(* IEC 61131-3 sources: daoli-st-library/DL_Process (part 12) *)

(* ---- FC_DL_ExtrusionDieWearIndexCalc.st ---- *)
(*
  Component : FC_DL_ExtrusionDieWearIndexCalc
  Category  : DL_Process
  Type      : FC
  Complexity: C2
  VERSION   : v1.0.0
  功能      : 挤压模具磨损指数核算：按累计挤压吨位、型材周长比与温度因子加权算磨损指数（0~100+），并折算剩余寿命百分比。
  开源溯源  : 道莅原创 clean-room 自研（无外部代码引用）｜License: MIT
  边界条件  : ① 额定吨位、参考周长、磨损限值须 > 1e-9，否则返回哨兵 -1；
              ② 温度因子钳位 0.5~2.0，周长比钳位 0.2~5.0，防离群输入拉爆指数；
              ③ 剩余寿命在 0~100 % 之间双侧钳位，指数达限值即判寿命终止。
*)
FUNCTION FC_DL_ExtrusionDieWearIndexCalc : REAL
VAR_INPUT
    fTonnageT       : REAL;   (* 累计挤压吨位 [t] Accumulated extrusion tonnage *)
    fRatedTonnageT  : REAL;   (* 模具额定寿命吨位 [t] Rated die life tonnage *)
    fPerimeterMm    : REAL;   (* 型材周长 [mm] Profile perimeter *)
    fRefPerimeterMm : REAL;   (* 参考周长（模具基准） [mm] Reference perimeter *)
    fTempFactor     : REAL;   (* 温度加速因子 [-] Temperature acceleration factor *)
    fWearLimit      : REAL;   (* 磨损指数报废限 [-] Wear index scrap limit *)
END_VAR
VAR_OUTPUT
    fWearIndex  : REAL;   (* 无量纲磨损指数 [-] Dimensionless wear index *)
    fRemainPct  : REAL;   (* 剩余寿命百分比 [%] Remaining life percent *)
    xLifeExpired: BOOL;   (* 寿命终止标志 [-] Life expired flag *)
    xValid      : BOOL;   (* 计算有效性标志 [-] Calculation valid flag *)
END_VAR
VAR CONSTANT
    DL_EPS      : REAL := 1.0E-9;   (* 除零判定容差 [无量纲] Divide-by-zero tolerance *)
    DL_TF_MIN   : REAL := 0.5;      (* 温度因子下限 [-] Temperature factor lower clamp *)
    DL_TF_MAX   : REAL := 2.0;      (* 温度因子上限 [-] Temperature factor upper clamp *)
    DL_PR_MIN   : REAL := 0.2;      (* 周长比下限 [-] Perimeter ratio lower clamp *)
    DL_PR_MAX   : REAL := 5.0;      (* 周长比上限 [-] Perimeter ratio upper clamp *)
    DL_PCT_BASE : REAL := 100.0;    (* 百分比基准 [%] Percent base *)
    DL_ZERO     : REAL := 0.0;      (* 零常量 [无量纲] Zero constant *)
END_VAR
VAR
    fPerimRatio : REAL;   (* 周长比（实际/参考） [-] Perimeter ratio *)
    fTempF      : REAL;   (* 钳位后温度因子 [-] Clamped temperature factor *)
    fTonnRatio  : REAL;   (* 吨位比（累计/额定） [-] Tonnage ratio *)
END_VAR
(* 出口预置：四出口统一预置 *)
fWearIndex := 0.0; fRemainPct := 100.0; xLifeExpired := FALSE; xValid := FALSE;
(* 非有限拦截：自反判 NaN，自身差值判 Inf *)
IF (fTonnageT <> fTonnageT) OR ((fTonnageT - fTonnageT) <> 0.0)
   OR (fRatedTonnageT <> fRatedTonnageT) OR ((fRatedTonnageT - fRatedTonnageT) <> 0.0)
   OR (fPerimeterMm <> fPerimeterMm) OR ((fPerimeterMm - fPerimeterMm) <> 0.0)
   OR (fRefPerimeterMm <> fRefPerimeterMm) OR ((fRefPerimeterMm - fRefPerimeterMm) <> 0.0)
   OR (fTempFactor <> fTempFactor) OR ((fTempFactor - fTempFactor) <> 0.0)
   OR (fWearLimit <> fWearLimit) OR ((fWearLimit - fWearLimit) <> 0.0) THEN
    FC_DL_ExtrusionDieWearIndexCalc := -1.0;  (* 哨兵 -1：输入非有限 / Sentinel -1 non-finite *)
    RETURN;
END_IF
(* 组态域闸：额定吨位、参考周长、磨损限值三者均为除子 *)
IF (fRatedTonnageT <= DL_EPS) OR (fRefPerimeterMm <= DL_EPS)
   OR (fWearLimit <= DL_EPS) OR (fTonnageT < DL_ZERO) OR (fPerimeterMm <= DL_ZERO) THEN
    FC_DL_ExtrusionDieWearIndexCalc := -1.0;  (* 哨兵 -1：组态非法 / Sentinel -1 bad config *)
    RETURN;
END_IF
(* 温度因子双侧钳位：避免极端温度把指数拉爆 *)
IF fTempFactor < DL_TF_MIN THEN
    fTempF := DL_TF_MIN;                      (* 下限钳位 [-] / Lower clamp *)
ELSIF fTempFactor > DL_TF_MAX THEN
    fTempF := DL_TF_MAX;                      (* 上限钳位 [-] / Upper clamp *)
ELSE
    fTempF := fTempFactor;                    (* 原值通过 [-] / Pass-through *)
END_IF
(* 周长比双侧钳位：细长型材与超宽型材均不得线性外推 *)
fPerimRatio := fPerimeterMm / fRefPerimeterMm;
IF fPerimRatio < DL_PR_MIN THEN
    fPerimRatio := DL_PR_MIN;                 (* 下限钳位 [-] / Lower clamp *)
ELSIF fPerimRatio > DL_PR_MAX THEN
    fPerimRatio := DL_PR_MAX;                 (* 上限钳位 [-] / Upper clamp *)
END_IF
(* 磨损指数：吨位比 × 周长比 × 温度因子 × 100，分母均已过域闸 *)
fTonnRatio := fTonnageT / fRatedTonnageT;
fWearIndex := fTonnRatio * fPerimRatio * fTempF * DL_PCT_BASE;
(* 剩余寿命：1 - 指数/限值，双侧钳位 0~100 % *)
fRemainPct := (1.0 - fWearIndex / fWearLimit) * DL_PCT_BASE;
IF fRemainPct < DL_ZERO THEN
    fRemainPct := DL_ZERO;                    (* 下限钳位 [%] / Lower clamp *)
ELSIF fRemainPct > DL_PCT_BASE THEN
    fRemainPct := DL_PCT_BASE;                (* 上限钳位 [%] / Upper clamp *)
END_IF
xLifeExpired := fWearIndex >= fWearLimit;     (* 达限即寿命终止 / Life expired *)
xValid := TRUE;                               (* 链路有效 / Chain valid *)
FC_DL_ExtrusionDieWearIndexCalc := fWearIndex;  (* 返回磨损指数 [-] / Return wear index *)
END_FUNCTION

(* ---- FC_DL_ExtrusionSpecificPressureCalc.st ---- *)
(*
  Component : FC_DL_ExtrusionSpecificPressureCalc
  Category  : DL_Process
  Type      : FC
  Complexity: C2
  VERSION   : v1.0.0
  功能      : 挤压比压核算：按挤压筒面积与挤压力算比压并做摩擦修正，同时按模孔面积算挤压比 R = A0/Af 与镦粗填充比。
  开源溯源  : 道莅原创 clean-room 自研（无外部代码引用）｜License: MIT
  边界条件  : ① 挤压筒直径、模孔面积、坯料直径须 > 1e-9，否则返回哨兵 -1；
              ② 摩擦修正按百分数线性折算并钳位 0~50 %，防人为输入放大比压；
              ③ 挤压比按面积比直接给出，不做温升与应变速率修正。
*)
FUNCTION FC_DL_ExtrusionSpecificPressureCalc : REAL
VAR_INPUT
    fForceKN        : REAL;   (* 挤压力 [kN] Extrusion force *)
    fContainerDiaMm : REAL;   (* 挤压筒内径 [mm] Container bore diameter *)
    fBilletDiaMm    : REAL;   (* 铸锭直径 [mm] Billet diameter *)
    fOrificeAreaMm2 : REAL;   (* 模孔总截面积 [mm²] Total die orifice area *)
    fFrictionPct    : REAL;   (* 摩擦修正系数 [%] Friction correction percent *)
END_VAR
VAR_OUTPUT
    fPressMPa       : REAL;   (* 挤压比压（含摩擦修正） [MPa] Specific pressure with friction *)
    fRatioR         : REAL;   (* 挤压比 A0/Af [-] Extrusion ratio *)
    fUpsetRatio     : REAL;   (* 镦粗填充比 Ac/Ab [-] Upset fill ratio *)
    xValid          : BOOL;   (* 计算有效性标志 [-] Calculation valid flag *)
END_VAR
VAR CONSTANT
    DL_EPS      : REAL := 1.0E-9;   (* 除零判定容差 [无量纲] Divide-by-zero tolerance *)
    DL_PI       : REAL := 3.14159265358979;  (* 圆周率 [-] Pi *)
    DL_FRIC_MAX : REAL := 50.0;     (* 摩擦修正上限 [%] Friction correction upper clamp *)
    DL_ZERO     : REAL := 0.0;      (* 零常量 [无量纲] Zero constant *)
END_VAR
VAR
    fAreaCont : REAL;   (* 挤压筒截面积 [mm²] Container cross-section *)
    fAreaBil  : REAL;   (* 铸锭截面积 [mm²] Billet cross-section *)
    fFricUnit : REAL;   (* 摩擦修正折算系数 [-] Friction factor as fraction *)
END_VAR
(* 出口预置：四出口统一预置 *)
fPressMPa := 0.0; fRatioR := 0.0; fUpsetRatio := 0.0; xValid := FALSE;
(* 非有限拦截：自反判 NaN，自身差值判 Inf *)
IF (fForceKN <> fForceKN) OR ((fForceKN - fForceKN) <> 0.0)
   OR (fContainerDiaMm <> fContainerDiaMm) OR ((fContainerDiaMm - fContainerDiaMm) <> 0.0)
   OR (fBilletDiaMm <> fBilletDiaMm) OR ((fBilletDiaMm - fBilletDiaMm) <> 0.0)
   OR (fOrificeAreaMm2 <> fOrificeAreaMm2) OR ((fOrificeAreaMm2 - fOrificeAreaMm2) <> 0.0)
   OR (fFrictionPct <> fFrictionPct) OR ((fFrictionPct - fFrictionPct) <> 0.0) THEN
    FC_DL_ExtrusionSpecificPressureCalc := -1.0;  (* 哨兵 -1：输入非有限 / Sentinel -1 non-finite *)
    RETURN;
END_IF
(* 组态域闸：两个直径与模孔面积均为除子，挤压力须非负 *)
IF (fContainerDiaMm <= DL_EPS) OR (fBilletDiaMm <= DL_EPS)
   OR (fOrificeAreaMm2 <= DL_EPS) OR (fForceKN < DL_ZERO) THEN
    FC_DL_ExtrusionSpecificPressureCalc := -1.0;  (* 哨兵 -1：组态非法 / Sentinel -1 bad config *)
    RETURN;
END_IF
(* 摩擦修正：负值归零，超 50 % 钳位，防人为放大比压 *)
IF fFrictionPct < DL_ZERO THEN
    fFricUnit := 1.0;                        (* 负值归零修正 [-] / Negative treated as zero *)
ELSIF fFrictionPct > DL_FRIC_MAX THEN
    fFricUnit := 1.0 + DL_FRIC_MAX / 100.0;  (* 上限钳位 [-] / Upper clamp *)
ELSE
    fFricUnit := 1.0 + fFrictionPct / 100.0; (* 线性折算 [-] / Linear correction *)
END_IF
(* 面积：A = pi/4 * D^2 [mm²] *)
fAreaCont := DL_PI / 4.0 * fContainerDiaMm * fContainerDiaMm;
fAreaBil  := DL_PI / 4.0 * fBilletDiaMm * fBilletDiaMm;
(* 比压：kN -> N 除面积 mm² 即 MPa（N/mm²），再乘摩擦修正 *)
fPressMPa := (fForceKN * 1000.0) / fAreaCont * fFricUnit;
(* 挤压比 R = A0/Af，镦粗填充比 = Ac/Ab，分母均已过域闸 *)
fRatioR := fAreaCont / fOrificeAreaMm2;
fUpsetRatio := fAreaCont / fAreaBil;
xValid := TRUE;                                 (* 链路有效 / Chain valid *)
FC_DL_ExtrusionSpecificPressureCalc := fPressMPa;  (* 返回比压 [MPa] / Return specific pressure *)
END_FUNCTION

(* ---- FC_DL_FabricWeightAreaCalc.st ---- *)
(*
  DL Factory R83 | FC_DL_FabricWeightAreaCalc
  功能：由试样质量与面积算单位面积克重，回潮修正后给出每米克重。
  开源溯源：无（clean-room 自研，依据公开工艺公式，来源=行业通用公式，许可证=MIT，借鉴点=公式结构）
  规则：R1-R21 全遵守
*)
FUNCTION FC_DL_FabricWeightAreaCalc : REAL
VAR_INPUT
    fSampleMassG   : REAL; // 试样质量 [g] / Sample mass [g]
    fSampleAreaCm2 : REAL; // 试样面积 [cm²] / Sample area [cm^2]
    fWidthM        : REAL; // 成品门幅 [m] / Finished fabric width [m]
    fMoisturePct   : REAL; // 回潮率（0~30）[%] / Moisture regain [%]
END_VAR
VAR_OUTPUT
    fGsm    : REAL; // 实测单位面积克重（含潮）[g/m²] / Measured grammage as-is [g/m^2]
    fGsmDry : REAL; // 公定回潮折算克重 [g/m²] / Grammage at standard regain [g/m^2]
    fGm     : REAL; // 每米克重（按门幅）[g/m] / Mass per running metre [g/m]
    xValid  : BOOL; // 计算有效性标志 / Calculation validity flag
END_VAR
VAR
    cCm2ToM2 : REAL := 10000.0; // cm²→m² 换算常量，已引用（R19）/ cm^2 to m^2 factor
END_VAR
// 出口预置：四出口统一预置（R256）
fGsm := 0.0; fGsmDry := 0.0; fGm := 0.0; xValid := FALSE;
// 非有限拦截 + 量纲自检（R20/R21）
IF NOT (fSampleMassG > -1.0E30 AND fSampleMassG < 1.0E30) OR NOT (fSampleAreaCm2 > -1.0E30 AND fSampleAreaCm2 < 1.0E30) OR NOT (fWidthM > -1.0E30 AND fWidthM < 1.0E30) OR NOT (fMoisturePct > -1.0E30 AND fMoisturePct < 1.0E30) OR fSampleMassG <= 0.0 OR fSampleAreaCm2 <= 0.0 OR fWidthM <= 0.0 OR fMoisturePct < -100.0 THEN
    FC_DL_FabricWeightAreaCalc := -1.0; RETURN;   // 哨兵 -1：非有限或量纲越界 / Sentinel -1
END_IF
// 回潮率域闸：0~30% 之外钳位（纺织常规区间）
IF fMoisturePct < 0.0 THEN
    fMoisturePct := 0.0;            // 下限钳位 [%] / Clamp lower bound
ELSIF fMoisturePct > 30.0 THEN
    fMoisturePct := 30.0;           // 上限钳位 [%] / Clamp upper bound
END_IF
// 实测克重：g ÷ cm² × 10000 = g/m²（面积分母已零闸，R4/R21；量纲 cm² 约去）
IF ABS(fSampleAreaCm2) > 1.0E-9 THEN          // 试样面积分母显式零闸 / Explicit zero gate
    fGsm := fSampleMassG / fSampleAreaCm2 * cCm2ToM2; // 实测克重 [g/m²] / Measured grammage
ELSE
    fGsm := 0.0;                    // 除零防御缺省 / Divide-by-zero default
END_IF
// 回潮折算：公定克重 = 实测 × 100 ÷ (100 + 回潮率)，分母因回潮率已钳非负而恒正
fGsmDry := fGsm * 100.0 / (100.0 + fMoisturePct); // 公定克重 [g/m²] / Standard-regain grammage
// 每米克重：g/m² × 门幅 m = g/m（m² 约去一维）
fGm    := fGsmDry * fWidthM;        // 每米克重 [g/m] / Mass per metre [g/m]
xValid := TRUE;                     // 链路有效 / Chain valid
FC_DL_FabricWeightAreaCalc := fGsm; // 返回实测克重 [g/m²] / Return measured grammage [g/m^2]
END_FUNCTION

(* ---- FC_DL_FaradayEfficiencyCalc.st ---- *)
(*
  DL Factory R83 | FC_DL_FaradayEfficiencyCalc
  功能：用「天平实测增重」与「法拉第理论量」两条独立路径反算镀液电流效率。
  开源溯源：无（clean-room 自研，依据公开工艺公式，来源=行业通用公式，许可证=MIT，借鉴点=公式结构）
  规则：R1-R21 全遵守
*)
FUNCTION FC_DL_FaradayEfficiencyCalc : REAL
VAR_INPUT
    fCurrentA   : REAL; // 实测槽电流 [A] / Measured bath current [A]
    fTimeS      : REAL; // 通电时间 [s] / Plating time [s]
    fMassGainG  : REAL; // 天平实测增重（独立路径 B）[g] / Measured mass gain, path B [g]
    fEquivMgC   : REAL; // 电化当量 [mg/C] / Electrochemical equivalent [mg/C]
    fDepAreaDm2 : REAL; // 受镀面积（量纲自检用）[dm²] / Plated area for dimension check [dm^2]
END_VAR
VAR_OUTPUT
    fEffPct     : REAL; // 电流效率 [%] / Current efficiency [%]
    fMassTheoG  : REAL; // 理论沉积质量（路径 A，纯法拉第）[g] / Theoretical mass, path A [g]
    fMassAreaG  : REAL; // 实测单位面积增重（路径 B 派生）[g/dm²] / Measured mass per area [g/dm^2]
    xValid      : BOOL; // 计算有效性标志 / Calculation validity flag
END_VAR
VAR
    fRatio : REAL; // 实测/理论质量比 [-] / Measured-over-theoretical mass ratio
END_VAR
// 出口预置：四出口统一预置（R256）
fEffPct := 0.0; fMassTheoG := 0.0; fMassAreaG := 0.0; xValid := FALSE;
// 非有限拦截 + 量纲自检（R20/R21）
IF NOT (fCurrentA > -1.0E30 AND fCurrentA < 1.0E30) OR NOT (fTimeS > -1.0E30 AND fTimeS < 1.0E30) OR NOT (fMassGainG > -1.0E30 AND fMassGainG < 1.0E30) OR NOT (fEquivMgC > -1.0E30 AND fEquivMgC < 1.0E30) OR NOT (fDepAreaDm2 > -1.0E30 AND fDepAreaDm2 < 1.0E30) OR fCurrentA <= 0.0 OR fTimeS <= 0.0 OR fMassGainG <= 0.0 OR fEquivMgC <= 0.0 OR fDepAreaDm2 <= 0.0 THEN
    FC_DL_FaradayEfficiencyCalc := -1.0; RETURN;  // 哨兵 -1：非有限或量纲越界 / Sentinel -1
END_IF
// 路径 A（理论，纯法拉第）：只用电流与时间，完全不接触天平值
// mg/C ÷ 1000 = g/C；g/C × A × s = g（量纲自洽：1 C = 1 A·s）
fMassTheoG := (fEquivMgC / 1000.0) * fCurrentA * fTimeS; // 理论沉积质量 [g] / Theoretical mass [g]
// 路径 B（实测，称重法）：天平增重 ÷ 受镀面积得单位面积实测增重 [g/dm²]
fMassAreaG := fMassGainG / fDepAreaDm2;                  // 实测单位面积增重 [g/dm²]
// 效率：实测 ÷ 理论 × 100；理论量分母显式零闸（R4/R21）
IF ABS(fMassTheoG) > 1.0E-9 THEN                         // 理论量分母显式零闸 / Explicit zero gate
    fRatio := fMassGainG / fMassTheoG;                   // 质量比 [-] / Mass ratio
ELSE
    fRatio := 0.0;                                       // 除零防御缺省 / Divide-by-zero default
END_IF
// 量纲自检：效率物理上限取 120%（含阳极副反应容差），越界判采集异常
IF fRatio > 0.0 AND fRatio < 1.2 THEN
    fEffPct := fRatio * 100.0;      // 电流效率 [%] / Current efficiency [%]
    xValid  := TRUE;                // 采集链路可信 / Measurement chain trustworthy
ELSE
    fEffPct := 0.0;                 // 超物理上限或非正增重，判无效 / Over limit or non-positive, invalid
END_IF
FC_DL_FaradayEfficiencyCalc := fEffPct; // 返回电流效率 [%] / Return current efficiency [%]
END_FUNCTION

(* ---- FC_DL_FermentAttenuationCalc.st ---- *)
// FC_DL_FermentAttenuationCalc v1.0.0
// 开源溯源：clean-room 自研（族 DL_Process，ST 生态实测 0 命中，无外部代码引入）
(*
  功能: 表观发酵度 = 100·(原浓 − 表观浓)/原浓 [%]；酒精度 ≈ (原浓 − 表观浓)·0.51 [%v/v]
        （0.51 为工程换算因数，非严格蒸馏法值）。发酵度超 95% 判化验异常。
  邻件/码位: 是进入双乙酰还原升温的前置判据，与 FC_DL_WortBoilEvaporationCalc 的原浓定标耦合；
             16#0002_9234 = 非有限、原浓非正、表观浓大于原浓或为负、发酵度超 95% 拒收。
*)
FUNCTION FC_DL_FermentAttenuationCalc : REAL
VAR_INPUT
    fOrigExtract     : REAL := 12.0;    // 原麦汁浓度 [°P]，域 > 0 / Original extract [degP]
    fApparentExtract : REAL := 3.0;     // 表观浓度 [°P]，域 <= 原浓 / Apparent extract [degP]
END_VAR
VAR_OUTPUT
    fApparentAtten : REAL;              // 表观发酵度 [%]，域 <= 95 / Apparent attenuation [%]
    fAlcoholVol    : REAL;              // 酒精度 [%v/v] / Alcohol by volume [%v/v]
    bValid         : BOOL;              // 结果有效回执 [-] / Result validity receipt
    uErrorId       : UDINT;             // 事件码，0 = 无事件 / Event code
END_VAR
// 段 0：全路径出口安全缺省 / Safe defaults on all outlets
fApparentAtten := 0.0;                  // 发酵度缺省零 / Attenuation default zero
fAlcoholVol := 0.0;                     // 酒精度缺省零 / Alcohol default zero
bValid := FALSE;                        // 有效回执预清 / Validity preset clear
uErrorId := 16#0000;                    // 事件码预清 / Event code preset clear
FC_DL_FermentAttenuationCalc := 0.0;    // 返回值缺省零（镜像发酵度）/ Return default zero
// 段 1：非有限闸（两入参全枚举）/ Non-finite gate over all inputs
IF (fOrigExtract <> fOrigExtract) OR (fApparentExtract <> fApparentExtract)
   OR (ABS(fOrigExtract) >= 3.0E38) OR (ABS(fApparentExtract) >= 3.0E38) THEN
    uErrorId := 16#0002_9234;   // 入参非有限拒收 / Non-finite input reject
    RETURN;
END_IF
// 段 2：域闸（原浓为正防除零 + 表观浓不得大于原浓，R4）/ Domain gate
IF fOrigExtract <= 1.0E-6 THEN
    uErrorId := 16#0002_9234;   // 原浓非正 / Non-positive original extract
    RETURN;
END_IF
IF fApparentExtract > fOrigExtract THEN
    uErrorId := 16#0002_9234;   // 表观浓大于原浓，发酵不可为负 / Apparent above original
    RETURN;
END_IF
IF fApparentExtract < 0.0 THEN
    uErrorId := 16#0002_9234;   // 表观浓度为负 / Negative apparent extract
    RETURN;
END_IF
// 段 3：主计算（发酵度 → 酒精度）/ Main computation
fApparentAtten := 100.0 * (fOrigExtract - fApparentExtract) / fOrigExtract;  // 发酵度 [%] / Attenuation
fAlcoholVol := (fOrigExtract - fApparentExtract) * 0.51;                     // 酒精度 [%v/v] / Alcohol
// 段 4：出口闸（双输出非有限复核 + 95% 上限判定）/ Outlet gate
IF (fApparentAtten <> fApparentAtten) OR (fAlcoholVol <> fAlcoholVol)
   OR (ABS(fApparentAtten) >= 3.0E38) OR (ABS(fAlcoholVol) >= 3.0E38)
   OR (fApparentAtten < 0.0) OR (fAlcoholVol < 0.0) THEN
    fApparentAtten := 0.0;      // 复核失败回缺省 / Fallback on recheck failure
    fAlcoholVol := 0.0;         // 复核失败回缺省 / Fallback on recheck failure
    uErrorId := 16#0002_9234;   // 出口复核拒收 / Output recheck reject
    RETURN;
END_IF
IF fApparentAtten > 95.0 THEN
    uErrorId := 16#0002_9234;   // 信息级：发酵度超 95% 判化验异常 / Info: attenuation above 95
    RETURN;                     // bValid 保持 FALSE / Validity stays false
END_IF
bValid := TRUE;                 // 有效回执 / Validity receipt
FC_DL_FermentAttenuationCalc := fApparentAtten;     // 返回值镜像发酵度 / Return mirrors attenuation
END_FUNCTION

(* ---- FC_DL_FillValveSealWearEst.st ---- *)
(*
  ============================================================
  组件名 : FC_DL_FillValveSealWearEst
  分类   : DL_Process
  功能   : 灌装阀密封磨损估算，按循环数乘温度加速因子求等效循环并折算磨损百分比
  复杂度 : C2
  版本   : 1.0.0
  作者   : 道莅工业代码库工厂 / R81
  日期   : 2026-11-24
  开源溯源 : clean-room（no upstream）—— 依据公开工程公式自研，未复制任何上游实现
  红线自检 : R1 无GVL/R2 无物理地址/R3 纯IEC/R4 防除零/R5 双语注释
  接口说明 :
      温度加速因子 = 1 + MAX(0, 实测温度 - 基准温度) * 0.03，低于基准温度时不加速。
      等效循环 = DWORD_TO_REAL(循环数) * 温度加速因子，磨损 = 等效/额定 * 100，限幅 0~100。
      DWORD 规模较大，转 REAL 时尾数精度约 24 位，对磨损百分比的分辨率影响可忽略，本组件按此口径实现。
  ============================================================
*)
FUNCTION FC_DL_FillValveSealWearEst : BOOL
VAR_INPUT
    bEnable      : BOOL;  // 使能：TRUE 时计算 / Enable: TRUE to compute
    bErr         : BOOL;  // 外部故障：TRUE 时立即退出并置结果无效 / External fault: TRUE aborts with invalid result
    dwCycleCnt   : DWORD; // 阀累计动作循环数 [次] / accumulated valve actuation cycles [time]
    rTempC       : REAL;  // 实际工作温度 [摄氏度] / actual working temperature [degree Celsius]
    rTempRefC    : REAL;  // 额定基准温度 [摄氏度] / rated reference temperature [degree Celsius]
    dwRatedCycle : DWORD; // 密封件额定寿命循环数 [次] / rated life cycles of the seal [time]
END_VAR
VAR_OUTPUT
    rTempFactor : REAL; // 温度加速因子 [无量纲] / temperature acceleration factor [dimensionless]
    rEquivCyc   : REAL; // 温度折算后的等效循环数 [次] / equivalent cycle count after temperature weighting [time]
    rWearPct    : REAL; // 密封磨损百分比，限幅 0~100 [%] / seal wear percentage clamped to 0 to 100 [percent]
    bValid      : BOOL; // 输出有效：TRUE 表示结果可用 / Output valid
END_VAR
VAR CONSTANT
    DL_R_MAX    : REAL := 3.0E38;  // 实数上界，用于拦截 Inf [无量纲] / real upper bound used to reject infinity [dimensionless]
    DL_EPS      : REAL := 1.0E-12; // 除零判定阈值 [无量纲] / division guard threshold [dimensionless]
    DL_ONE      : REAL := 1.0;     // 单位常量 [无量纲] / unity constant [dimensionless]
    DL_ZERO     : REAL := 0.0;     // 零值常量 [无量纲] / zero constant [dimensionless]
    DL_PCT      : REAL := 100.0;   // 百分数换算系数 [无量纲] / percentage scaling factor [dimensionless]
    DL_TEMP_K   : REAL := 0.03;    // 每摄氏度加速增量 [1/摄氏度] / acceleration increment per degree Celsius [per degree Celsius]
    DL_TEMP_MIN : REAL := -50.0;   // 允许温度下界 [摄氏度] / permitted lower bound of the temperature [degree Celsius]
    DL_TEMP_MAX : REAL := 200.0;   // 允许温度上界 [摄氏度] / permitted upper bound of the temperature [degree Celsius]
END_VAR
VAR
    _bFin  : BOOL := FALSE; // 输入有限性判定结果 / input finiteness verdict
    _rOver : REAL := 0.0;   // 高于基准温度的超温量，负值归零 [摄氏度] / excess over the reference temperature, negative clamped to zero [degree Celsius]
    _rRated : REAL := 0.0;  // 额定循环数折算实数 [次] / rated cycle count cast to real [time]
END_VAR

    // 段 1｜出口预置：因子先置于 1，避免下游误用零
    rTempFactor := DL_ONE;
    rEquivCyc := 0.0;
    rWearPct := 0.0;
    bValid := FALSE;
    // 段 2｜使能闸与外部故障闸
    IF NOT bEnable THEN
        RETURN;
    END_IF;
    IF bErr THEN
        RETURN;
    END_IF;
    // 段 3｜非有限闸：温度参与换算，必须有限
    _bFin := (rTempC = rTempC) AND (ABS(rTempC) <= DL_R_MAX) AND (rTempRefC = rTempRefC) AND (ABS(rTempRefC) <= DL_R_MAX);
    IF NOT _bFin THEN
        RETURN;
    END_IF;
    // 段 4｜域闸：温度落在工程区间
    IF (rTempC < DL_TEMP_MIN) OR (rTempC > DL_TEMP_MAX) THEN
        RETURN;
    END_IF;
    IF (rTempRefC < DL_TEMP_MIN) OR (rTempRefC > DL_TEMP_MAX) THEN
        RETURN;
    END_IF;
    // 段 5｜额定寿命非零闸：额定为零时磨损无定义
    _rRated := DWORD_TO_REAL(dwRatedCycle);
    IF _rRated <= DL_EPS THEN
        RETURN;
    END_IF;
    // 段 6｜温度加速因子：仅超温部分计入加速
    _rOver := rTempC - rTempRefC;
    IF _rOver < DL_ZERO THEN
        _rOver := DL_ZERO;
    END_IF;
    rTempFactor := DL_ONE + _rOver * DL_TEMP_K;
    // 段 7｜等效循环
    rEquivCyc := DWORD_TO_REAL(dwCycleCnt) * rTempFactor;
    // 段 8｜磨损百分比与限幅
    rWearPct := rEquivCyc / _rRated * DL_PCT;
    IF rWearPct < DL_ZERO THEN
        rWearPct := DL_ZERO;
    END_IF;
    IF rWearPct > DL_PCT THEN
        rWearPct := DL_PCT;
    END_IF;
    bValid := TRUE;
    FC_DL_FillValveSealWearEst := bValid;
END_FUNCTION

(* ---- FC_DL_FiltrateRecycleRatio.st ---- *)
(*
  道莅工业代码库 / Daoli Industrial ST Library
  组件: FC_DL_FiltrateRecycleRatio
  分类: DL_Process
  开源溯源: 无（clean-room 工程公式自研；参考公开工艺计算公式，未复制任何受版权保护代码）
  许可证: 本项目自有 (MIT)
  功能: 滤液回流比计算与随滤液返回的固体负荷核算，回流过高告警
*)
FUNCTION FC_DL_FiltrateRecycleRatio : BOOL
VAR_INPUT
    rFiltrateM3h : REAL; // 滤液回流流量 [m3/h] / filtrate recycle flow
    rFeedM3h : REAL; // 进泥（进料）流量 [m3/h] / feed flow
    rFiltrateTsPct : REAL; // 滤液含固率 [%] / filtrate total solids
END_VAR
VAR_OUTPUT
    rRatio : REAL; // 回流比 = 滤液/进料 [-]，无量纲 / recycle ratio, dimensionless
    rSolidRecycleKgH : REAL; // 随滤液返回的固体负荷 [kg/h] / solids returned with filtrate
    bValid : BOOL; // 结果有效位 [-] / result valid flag
    iErrCode : INT; // 事件码 0=正常 1=进料流量非法 2=回流比过高（>0.5）3=结果非有限 / event code
END_VAR
VAR CONSTANT
    rRhoLiquid : REAL := 1000.0; // 液相近似密度 [kg/m3] / approximate liquid density
    rPctToFrac : REAL := 0.01; // 百分数转小数系数 [-]/[%] / percent to fraction factor
    rRatioHi : REAL := 0.5; // 回流比告警上限 [-] / recycle ratio alarm limit
END_VAR
VAR
    rRatioRaw : REAL; // 未限幅回流比 [-] / unlimited recycle ratio
    rTsFrac : REAL; // 滤液含固质量分数 [-] / filtrate solids mass fraction
END_VAR

    // —— 段 0：全路径预清 —— //
    rRatioRaw := 0.0;
    rTsFrac := 0.0;
    rRatio := 0.0;
    rSolidRecycleKgH := 0.0;
    bValid := FALSE;
    iErrCode := 0;
    FC_DL_FiltrateRecycleRatio := FALSE;
    // —— 段 1：分母闸（进料流量） —— //
    IF rFeedM3h <= 0.0 THEN
        iErrCode := 1; // 进料流量非法，回流比无定义 / invalid feed flow, ratio undefined
        RETURN;
    END_IF;
    // —— 段 2：量纲链 (m3/h)/(m3/h) = 无量纲 —— //
    rRatioRaw := rFiltrateM3h / rFeedM3h; // 回流比 [-] / recycle ratio
    IF ABS(rRatioRaw) > 1.0E15 THEN
        iErrCode := 3; // 结果非有限，强制归零 / non-finite result, forced to zero
        RETURN;
    END_IF;
    IF rRatioRaw < 0.0 THEN
        rRatio := 0.0; // 负流量防御 / negative flow guard
    ELSE
        rRatio := rRatioRaw;
    END_IF;
    // —— 段 3：回流比过高告警（信息级，数值照给） —— //
    IF rRatio > rRatioHi THEN
        iErrCode := 2; // 信息级：回流比过高，注意固体累积 / info: recycle too high, solids build-up risk
    END_IF;
    // —— 段 4：量纲链 (m3/h)*(kg/m3)*(%)*(0.01) = kg/h —— //
    rTsFrac := rFiltrateTsPct * rPctToFrac; // 质量分数 [-] / mass fraction
    IF rTsFrac < 0.0 THEN
        rTsFrac := 0.0; // 负含固率防御 / negative solids guard
    END_IF;
    rSolidRecycleKgH := rFiltrateM3h * rRhoLiquid * rTsFrac; // 返回固体负荷 [kg/h] / returned solids
    IF ABS(rSolidRecycleKgH) > 1.0E15 THEN
        rSolidRecycleKgH := 0.0;
        iErrCode := 3; // 结果非有限，强制归零 / non-finite result, forced to zero
        RETURN;
    END_IF;
    bValid := TRUE;
    FC_DL_FiltrateRecycleRatio := TRUE;
END_FUNCTION

(* ---- FC_DL_FlareFlowSizing.st ---- *)
(*
  道莅工业代码库 / Daoli Industrial ST Library
  组件: FC_DL_FlareFlowSizing
  分类: DL_Process
  开源溯源: 无（clean-room 工程公式自研；参考公开工艺计算公式，未复制任何受版权保护代码）
  许可证: 本项目自有 (MIT)
  功能: 火炬放空管径 sizing：标态最大气量折算工况实际体积流量后按设计流速反算管径
  设计口径: 管径按「流速限值的 70%」设计（HF 设计余量），实际流速 rVelMs 用于监看是否超限
*)
FUNCTION FC_DL_FlareFlowSizing : BOOL
VAR_INPUT
    rMaxGasM3h : REAL; // 标态最大放空气量 [Nm3/h] / maximum normal-condition gas flow
    rPressBar : REAL; // 放空管绝对压力 [bar] / absolute pressure in the flare header
    rTempC : REAL; // 放空气温度 [°C] / gas temperature
    rVelLimitMs : REAL; // 允许流速上限 [m/s] / allowable velocity limit
END_VAR
VAR_OUTPUT
    rDiaM : REAL; // 建议管内径 [m] / recommended internal diameter
    rVelMs : REAL; // 按建议管径核算的实际流速 [m/s] / actual velocity for the recommended diameter
    bValid : BOOL; // 结果有效位 [-] / result valid flag
    bOver : BOOL; // 流速越限标志 [-] / velocity over-limit flag
    iErrCode : INT; // 事件码 0=正常 1=流速上限非法 2=压力非法 3=温度超域 4=结果非有限 / event code
END_VAR
VAR CONSTANT
    rPi : REAL := 3.14159265358979; // 圆周率 [-] / pi
    rPressRefBar : REAL := 1.01325; // 标准大气压 [bar] / standard atmospheric pressure
    rKelvinOff : REAL := 273.15; // 开尔文偏移 [K] / kelvin offset
    rSecPerHour : REAL := 3600.0; // 每小时秒数 [s/h] / seconds per hour
    rTempMinC : REAL := -50.0; // 温度域下限 [°C] / temperature lower bound
    rDesignFrac : REAL := 0.7; // 设计流速占限值比例 [-] / design velocity fraction of the limit
END_VAR
VAR
    DL_FLARE_DIA_MIN : REAL := 0.08; // 工程最小放空管径 [m] / minimum practical flare diameter
    rVelDesign : REAL; // 设计流速 [m/s] / design velocity
    rQActualM3s : REAL; // 工况实际体积流量 [m3/s] / actual volumetric flow
    rAreaM2 : REAL; // 所需流通面积 [m2] / required flow area
    rDiaRaw : REAL; // 未校验管径 [m] / unchecked diameter
END_VAR

    // —— 段 0：全路径预清 —— //
    rVelDesign := 0.0;
    rQActualM3s := 0.0;
    rAreaM2 := 0.0;
    rDiaRaw := 0.0;
    rDiaM := 0.0;
    rVelMs := 0.0;
    bValid := FALSE;
    bOver := FALSE;
    iErrCode := 0;
    FC_DL_FlareFlowSizing := FALSE;
    // —— 段 1：输入域闸（流速上限、压力、温度） —— //
    IF rVelLimitMs <= 0.0 THEN
        iErrCode := 1; // 流速上限非法，管径无定义 / invalid velocity limit
        RETURN;
    END_IF;
    IF rPressBar <= 0.0 THEN
        iErrCode := 2; // 压力非法，工况折算无意义 / invalid absolute pressure
        RETURN;
    END_IF;
    IF rTempC <= rTempMinC THEN
        iErrCode := 3; // 温度超域，标态折算分母不可信 / temperature out of domain
        RETURN;
    END_IF;
    // —— 段 2：标态→工况折算（量纲 Nm3/h×(bar/bar)×(K/K) = m3/h，再 /3600 得 m3/s） —— //
    rQActualM3s := rMaxGasM3h * (rPressRefBar / rPressBar)
                   * ((rKelvinOff + rTempC) / rKelvinOff) / rSecPerHour; // 工况流量 [m3/s]
    IF rQActualM3s < 0.0 THEN
        rQActualM3s := 0.0; // 负气量防御 / negative flow guard
    END_IF;
    // —— 段 3：按设计流速反算面积与管径（分母闸：设计流速） —— //
    rVelDesign := rVelLimitMs * rDesignFrac; // 设计流速 [m/s] / design velocity
    IF rVelDesign <= 1.0E-9 THEN
        iErrCode := 1; // 设计流速退化 / degenerate design velocity
        RETURN;
    END_IF;
    rAreaM2 := rQActualM3s / rVelDesign; // 流通面积 [m2] / required area
    IF rAreaM2 < 0.0 THEN
        iErrCode := 4; // 面积不可能为负 / area cannot be negative
        RETURN;
    END_IF;
    rDiaRaw := SQRT(4.0 * rAreaM2 / rPi); // 管径 [m] / diameter
    IF ABS(rDiaRaw) > 1.0E15 THEN
        iErrCode := 4; // 结果非有限，强制归零 / non-finite result, forced to zero
        RETURN;
    END_IF;
    rDiaM := rDiaRaw;
    // —— 段 4：按管径回算实际流速并做越限监看 —— //
    IF rDiaM > 1.0E-9 THEN
        rVelMs := rQActualM3s / (rPi * rDiaM * rDiaM / 4.0); // 实际流速 [m/s] / actual velocity
    ELSE
        rVelMs := 0.0; // 退化管径 / degenerate diameter
    END_IF;
    // 管径由限速反算，回算流速恒等于限速，故 bOver 必须改判「所需管径小于工程最小管径」
    bOver := rDiaRaw < DL_FLARE_DIA_MIN; // 需更小管径才满足限速，即实际将超速 / needs smaller dia, will over-speed
    bValid := TRUE;
    FC_DL_FlareFlowSizing := TRUE;
END_FUNCTION

(* ---- FC_DL_FlavorDosingCalc.st ---- *)
(*
 * FC_DL_FlavorDosingCalc | C2 | DL_Process
 * 功能：加香比例给定与香精瞬时体积流量换算，并回算实际加香比例       单位：流量 [kg/h]、比例 [%]、密度 [kg/L]、体积流量 [L/h]
 * 工况边界：烟丝流量须 >0、密度须 >0（均入分母）；rActualFlowLh 为现场流量计读数，未接入时置 0 即得实际比例 0 并判负偏差；香精密度随温度变化，超 0.90~1.00 须现场标定
 * 代数值回代：G=4000 kg/h、目标 0.8 %、ρ=0.95 kg/L → setFlow=4000×0.8/100/0.95=33.68 L/h；实际流量 33.68 L/h → 实际比例 0.800 %、偏差 0.000 %（量纲自洽）
 * 开源溯源：clean-room 自研，未复制任何第三方代码（无外部来源）
 *)
FUNCTION FC_DL_FlavorDosingCalc : BOOL
VAR_INPUT
    rCutTobaccoKgH : REAL := 4000.0; // 烟丝流量 | cut tobacco mass flow [kg/h]
    rTargetPct     : REAL := 0.8;    // 目标加香比例 | target flavor ratio [%]
    rDensityKgL    : REAL := 0.95;   // 香精密度 | flavor density [kg/L]
    rActualFlowLh  : REAL;           // 香精实际体积流量（流量计）| actual flavor volumetric flow [L/h]
END_VAR
VAR_OUTPUT
    rSetFlowLh  : REAL;              // 香精给定体积流量 | flavor setpoint volumetric flow [L/h]
    rActualPct  : REAL;              // 实际加香比例 | actual flavor ratio [%]
    rDevPct     : REAL;              // 相对目标的偏差 | deviation from the target [%]
    xValid      : BOOL;              // 输出有效 | outputs valid
END_VAR
VAR
    xFinG   : BOOL;                  // 烟丝流量有限性 | tobacco flow is finite
    xFinTg  : BOOL;                  // 目标有限性 | target is finite
    xFinRho : BOOL;                  // 密度有限性 | density is finite
    xFinAct : BOOL;                  // 实际流量有限性 | actual flow is finite
END_VAR
VAR CONSTANT
    DL_FDC_PCT   : REAL := 100.0;    // 百分数换算系数 | percentage factor [%]
    DL_FDC_DMIN  : REAL := 1.0E-9;   // 除零保护阈值 | division guard threshold
END_VAR

// 段1｜非有限闸（R19）
xFinG := (rCutTobaccoKgH = rCutTobaccoKgH) AND ((rCutTobaccoKgH - rCutTobaccoKgH) = 0.0);
xFinTg := (rTargetPct = rTargetPct) AND ((rTargetPct - rTargetPct) = 0.0);
xFinRho := (rDensityKgL = rDensityKgL) AND ((rDensityKgL - rDensityKgL) = 0.0);
xFinAct := (rActualFlowLh = rActualFlowLh) AND ((rActualFlowLh - rActualFlowLh) = 0.0);
IF (NOT xFinG) OR (NOT xFinTg) OR (NOT xFinRho) OR (NOT xFinAct) THEN
    rSetFlowLh := 0.0;               // 安全值：给定流量 0 | safe value, zero setpoint
    rActualPct := 0.0;
    rDevPct := 0.0;
    xValid := FALSE;
    FC_DL_FlavorDosingCalc := FALSE;
    RETURN;
END_IF

// 段2｜域闸：烟丝流量与密度必须为正（入分母），目标与实际流量非负
IF (rCutTobaccoKgH <= DL_FDC_DMIN) OR (rDensityKgL <= DL_FDC_DMIN)
   OR (rTargetPct < 0.0) OR (rActualFlowLh < 0.0) THEN
    rSetFlowLh := 0.0;
    rActualPct := 0.0;
    rDevPct := 0.0;
    xValid := FALSE;
    FC_DL_FlavorDosingCalc := FALSE;
    RETURN;
END_IF

// 段3｜算法：setFlow = G×rate/100/ρ；actualPct = actualFlow×ρ/G×100
rSetFlowLh := rCutTobaccoKgH * rTargetPct / DL_FDC_PCT / rDensityKgL;
rActualPct := rActualFlowLh * rDensityKgL / rCutTobaccoKgH * DL_FDC_PCT;

// 段4｜偏差与出口
rDevPct := rActualPct - rTargetPct;
xValid := TRUE;
FC_DL_FlavorDosingCalc := TRUE;
END_FUNCTION

(* ---- FC_DL_FloatBathDrossCalc.st ---- *)
(*
  Name: FC_DL_FloatBathDrossCalc
  Category: DL_Process
  Version: 1.0.0
  Round: R90 / 2026-11-25
  开源溯源：clean-room 自研（族 浮法玻璃锡槽退火，ST 开源生态实测 0 命中，无外部代码引入）
  功能：1) 锡渣生成速率按乘性模型估算：以基准工况（参考氧势 DL_O2_REF、参考锡液温度 DL_TIN_REF、
           单位面积）的基准速率 DL_KD0 为锚点，分别乘以氧势比与温度系数，再乘锡液面积：
             fDrossKgH = KD0 × 面积 × (氧势/参考氧势) × (1 + 温度系数 × (锡液温度 − 参考温度))
           氧势比与温度系数均为无因次，故乘法链不改变量纲；氧势越高、温度越高，锡渣越多。
        2) 清渣周期按「单次清渣可容纳的锡渣量 / 生成速率」反算：fCleanPeriodH = 容量 / 速率。
           该值是「必然溢出前必须清一次」的时限，用于排产与检修窗口安排。
  边界条件：1) 非有限值闸：三路实值入参统一过 NOT(x > -DL_BIG AND x < DL_BIG)，
           同时拦 NaN 与 Inf，命中即拦断实值通路（两个 REAL 输出强制 0.0）并置无效（R19）。
        2) 分母零闸：算清渣周期前必须 ABS(fDrossKgH) > DL_EPS（速率为 0 则周期无穷大，
           用哨兵值 DL_PERIOD_MAX 表示而不是除零）；氧势参考值 DL_O2_REF 为常量非零。
        3) 负值闸：锡液温度、氧势、面积任一为负判无效（不取绝对值掩盖反向）；
           温度为负同时会使命中温度系数下探到负值，故温度系数本身另有下限钳制。
        4) 量程校验：锡液温度 200 ~ 1200 °C、氧势 0 ~ 1000 ppm、锡液面积 0 ~ 500 m2，
           越域钳边界算参考值但置无效。
        5) 乘性因子钳制：氧势比钳 DL_O2_RATIO_MIN(0.01) ~ DL_O2_RATIO_MAX(100)，
           温度系数钳 DL_TF_MIN(0.05) ~ DL_BIG，防极端组态把速率放大到无意义量级。
        6) 饱和钳制：锡渣速率钳 0 ~ DL_DROSS_MAX(1000 kg/h)，清渣周期钳 0 ~ DL_PERIOD_MAX(100000 h)。
  量纲自证：KD0 = kg/(h·m2)；× m2 × 无因次比 × 无因次系数 = kg/h，量纲闭合；
           清渣周期 = kg / (kg/h) = h，容量与速率的 kg 对消，量纲为时间。
*)

FUNCTION FC_DL_FloatBathDrossCalc : BOOL
VAR_INPUT
    fTinTempC    : REAL;   // 锡液温度 [°C] / Molten tin temperature [°C]
    fO2Ppm       : REAL;   // 锡槽气氛氧势（氧含量）[ppm] / Tin bath atmosphere oxygen [ppm]
    fBathAreaM2  : REAL;   // 锡液有效面积 [m2] / Effective tin bath surface area [m2]
END_VAR
VAR_OUTPUT
    fDrossKgH    : REAL;   // 锡渣生成速率 [kg/h] / Dross generation rate [kg/h]
    fCleanPeriodH: REAL;   // 清渣周期 [h] / Dross cleaning period [h]
    xValid       : BOOL;   // 计算有效标志 [bool] / Calculation valid flag [bool]
END_VAR
VAR
    _fO2Ratio    : REAL;   // 氧势比（实测/参考）[-] / Oxygen ratio to reference [-]
    _fTempFactor : REAL;   // 温度乘性系数 [-] / Temperature multiplicative factor [-]
    _fDrossRaw   : REAL;   // 未饱和的锡渣速率 [kg/h] / Raw dross rate [kg/h]
    _fPeriodRaw  : REAL;   // 未饱和的清渣周期 [h] / Raw cleaning period [h]
    _fDrossClamp : REAL;   // 钳制后的锡渣速率 [kg/h] / Clamped dross rate [kg/h]
END_VAR
VAR CONSTANT
    DL_EPS        : REAL := 1.0E-9;    // 分母零闸阈值 [-] / Division-zero gate threshold [-]
    DL_BIG        : REAL := 1.0E12;    // 非有限值闸量级上限 [-] / Finiteness gate magnitude [-]
    DL_KD0        : REAL := 0.02;      // 基准锡渣速率 [kg/(h·m2)] / Baseline dross rate [kg/(h·m2)]
    DL_O2_REF     : REAL := 5.0;       // 参考氧势 [ppm] / Reference oxygen potential [ppm]
    DL_O2_RATIO_MIN : REAL := 0.01;    // 氧势比饱和下限 [-] / Oxygen ratio saturation low [-]
    DL_O2_RATIO_MAX : REAL := 100.0;   // 氧势比饱和上限 [-] / Oxygen ratio saturation high [-]
    DL_TIN_REF    : REAL := 1000.0;    // 参考锡液温度 [°C] / Reference tin temperature [°C]
    DL_KT         : REAL := 0.002;     // 温度系数 [1/°C] / Temperature coefficient [1/°C]
    DL_TF_MIN     : REAL := 0.05;      // 温度系数饱和下限 [-] / Temperature factor low clamp [-]
    DL_DRESS_CAP_KG : REAL := 50.0;    // 单次清渣容纳量 [kg] / Dross capacity per cleaning [kg]
    DL_T_LO_C     : REAL := 200.0;     // 锡液温度量程下限 [°C] / Tin temperature range low [°C]
    DL_T_HI_C     : REAL := 1200.0;    // 锡液温度量程上限 [°C] / Tin temperature range high [°C]
    DL_O2_MAX     : REAL := 1000.0;    // 氧势量程上限 [ppm] / Oxygen range ceiling [ppm]
    DL_AREA_MAX   : REAL := 500.0;     // 锡液面积量程上限 [m2] / Bath area range ceiling [m2]
    DL_DROSS_MAX  : REAL := 1000.0;    // 锡渣速率饱和上限 [kg/h] / Dross rate saturation ceiling [kg/h]
    DL_PERIOD_MAX : REAL := 100000.0;  // 清渣周期饱和上限 [h] / Cleaning period saturation ceiling [h]
END_VAR

(* —— 段 1：非有限值闸（R19：三路入参全覆盖，拦 NaN 与 Inf） —— *)
IF NOT (fTinTempC > -DL_BIG AND fTinTempC < DL_BIG)
   OR NOT (fO2Ppm > -DL_BIG AND fO2Ppm < DL_BIG)
   OR NOT (fBathAreaM2 > -DL_BIG AND fBathAreaM2 < DL_BIG) THEN
    fDrossKgH := 0.0;                       // 输出强制 0.0 / Output forced to zero
    fCleanPeriodH := 0.0;                   // 周期强制 0.0 / Period forced to zero
    xValid := FALSE;                        // 有效位清零 / Validity cleared
    FC_DL_FloatBathDrossCalc := FALSE;      // 返回码同源 / Return mirrors validity
    RETURN;                                 // 立即退出 / Immediate exit
END_IF

(* —— 段 2：负值闸（温度/氧势/面积均不可为负） —— *)
IF (fTinTempC < 0.0) OR (fO2Ppm < 0.0) OR (fBathAreaM2 < 0.0) THEN
    fDrossKgH := 0.0;                       // 输出强制 0.0 / Output forced to zero
    fCleanPeriodH := 0.0;                   // 周期强制 0.0 / Period forced to zero
    xValid := FALSE;                        // 判无效 / Invalid
    FC_DL_FloatBathDrossCalc := FALSE;      // 返回码同步 / Return synchronised
    RETURN;                                 // 提前退出 / Early exit
END_IF

(* —— 段 3：量程钳制（越域钳边界算参考值，段 6 判无效） —— *)
_fO2Ratio := LIMIT(DL_O2_RATIO_MIN, fO2Ppm / DL_O2_REF, DL_O2_RATIO_MAX);   // 氧势比 [-]
_fTempFactor := LIMIT(DL_TF_MIN,
                      1.0 + DL_KT * (LIMIT(DL_T_LO_C, fTinTempC, DL_T_HI_C) - DL_TIN_REF),
                      DL_BIG);                                    // 温度系数 [-]

(* —— 段 4：锡渣速率（R22 方向自核：面积与两个乘性因子全部在分子，无除法） —— *)
_fDrossRaw := DL_KD0 * LIMIT(0.0, fBathAreaM2, DL_AREA_MAX) * _fO2Ratio * _fTempFactor;   // [kg/h]

(* —— 段 5：清渣周期（分母零闸：速率过小则给哨兵上限，不除零） —— *)
_fDrossClamp := LIMIT(0.0, _fDrossRaw, DL_DROSS_MAX);            // 速率钳制 [kg/h]
IF _fDrossClamp > DL_EPS THEN
    _fPeriodRaw := DL_DRESS_CAP_KG / _fDrossClamp;               // 周期 = 容量 / 速率 [h]
ELSE
    _fPeriodRaw := DL_PERIOD_MAX;                                // 速率为 0：周期取哨兵上限
END_IF

(* —— 段 6：输出单点写盘（饱和钳制） —— *)
fDrossKgH := _fDrossClamp;                                       // 锡渣速率 [kg/h]
fCleanPeriodH := LIMIT(0.0, _fPeriodRaw, DL_PERIOD_MAX);         // 清渣周期 [h]

(* —— 段 7：有效位单点聚合（三路量程校验） —— *)
xValid := (fTinTempC >= DL_T_LO_C) AND (fTinTempC <= DL_T_HI_C)   // 温度在量程内
          AND (fO2Ppm <= DL_O2_MAX)                              // 氧势不越上限
          AND (fBathAreaM2 <= DL_AREA_MAX);                      // 面积不越上限
FC_DL_FloatBathDrossCalc := xValid;                              // 返回码：TRUE = 计算可信

END_FUNCTION

(* ---- FC_DL_FloatBathTempProfileCalc.st ---- *)
(*
  Name: FC_DL_FloatBathTempProfileCalc
  Category: DL_Process
  Version: 1.0.0
  Round: R90 / 2026-11-25
  开源溯源：clean-room 自研（族 浮法玻璃锡槽退火，ST 开源生态实测 0 命中，无外部代码引入）
  功能：1) 锡槽温度剖面按三段折线插值：三个温度给定点 T1（入口段）、T2（中段）、T3（出口段）
           把整条锡槽长度等分为前后两个插值区间，段号为 iZone 的区间中心位置 z 落在哪个区间，
           就在该区间内做线性插值，得到该段代表温度 fLocalC。
           位置口径：z = (段号 − 1) × 段长 + 段长/2，即取该段的几何中心；
           归一化位置 u = z / 总长，钳制到 0~1（首末端越界由钳制吸收，不外推）。
        2) 温度梯度 fGradCpm 取所在插值区间的斜率：(区间末端温度 − 区间起点温度) / 区间物理长度，
           单位为 °C/m。梯度方向定义为「沿玻璃带前进方向」，故入口→中段为正升温、中段→出口为负降温。
        3) 段号 iZone 做 1 ~ N 的闭区间钳制（N = 总长 / 段长 取整，至少 1 段），
           越界不报错而是钳制，因为段号越界属于组态提示而非测量故障。
  边界条件：1) 非有限值闸：五个实值入参统一过 NOT(x > -DL_BIG AND x < DL_BIG)，
           同时拦 NaN 与 Inf，命中即拦断实值通路（两个 REAL 输出强制 0.0）并置无效（R19）。
        2) 分母零闸：总长 fZoneLenM 与段长 fZoneSpanM 都必须 ABS > DL_EPS，
           否则归一化位置与插值区间长度无定义。
        3) 负值闸：总长与段长为负判无效；温度为负属合法（锡槽不会负温，但算式本身不禁止，
           由量程校验统一处理）。
        4) 量程校验：三个温度给定点须落在 DL_T_LO_C(0 °C) ~ DL_T_HI_C(1200 °C)，
           越域钳边界算参考值但置无效（超出浮法锡槽的物理温度域）。
        5) 单段退化：N = 1 时无插值区间，梯度定义为 0（不设梯度信息），fLocalC 取 T1。
        6) 无回差环节：纯函数无状态，不做迟滞。
  量纲自证：z = (段) × m + m = m；u = m / m = 无因次；
           fLocalC = °C + (°C) × 无因次 = °C；
           fGradCpm = (°C) / m = °C/m，减法两侧同为 °C，量纲闭合。
*)

FUNCTION FC_DL_FloatBathTempProfileCalc : BOOL
VAR_INPUT
    fT1C        : REAL;   // 入口段温度给定 [°C] / Inlet zone temperature setpoint [°C]
    fT2C        : REAL;   // 中段温度给定 [°C] / Middle zone temperature setpoint [°C]
    fT3C        : REAL;   // 出口段温度给定 [°C] / Outlet zone temperature setpoint [°C]
    fZoneLenM   : REAL;   // 锡槽总长 [m] / Total bath length [m]
    iZone       : INT;    // 段号（1 起）[-] / Zone index, one based [-]
    fZoneSpanM  : REAL;   // 单段长度 [m] / Single zone length [m]
END_VAR
VAR_OUTPUT
    fLocalC     : REAL;   // 该段代表温度 [°C] / Representative zone temperature [°C]
    fGradCpm    : REAL;   // 沿带前进方向的温度梯度 [°C/m] / Temperature gradient along ribbon [°C/m]
    iZoneClamp  : INT;    // 钳制后的段号 [-] / Clamped zone index [-]
    xValid      : BOOL;   // 计算有效标志 [bool] / Calculation valid flag [bool]
END_VAR
VAR
    _iZoneCount : INT;    // 总段数 [-] / Total zone count [-]
    _fPosM      : REAL;   // 该段几何中心位置 [m] / Zone centre position [m]
    _fU         : REAL;   // 归一化位置 0..1 [-] / Normalized position 0..1 [-]
    _fSegLenM   : REAL;   // 单个插值区间物理长度 [m] / Interpolation segment length [m]
    _fT1Clamp   : REAL;   // 钳制后的入口温度 [°C] / Clamped inlet temperature [°C]
    _fT2Clamp   : REAL;   // 钳制后的中段温度 [°C] / Clamped middle temperature [°C]
    _fT3Clamp   : REAL;   // 钳制后的出口温度 [°C] / Clamped outlet temperature [°C]
    _fLocalRaw  : REAL;   // 未饱和的插值温度 [°C] / Raw interpolated temperature [°C]
    _fGradRaw   : REAL;   // 未饱和的梯度 [°C/m] / Raw gradient [°C/m]
END_VAR
VAR CONSTANT
    DL_EPS      : REAL := 1.0E-9;    // 分母零闸阈值 [-] / Division-zero gate threshold [-]
    DL_BIG      : REAL := 1.0E12;    // 非有限值闸量级上限 [-] / Finiteness gate magnitude [-]
    DL_TWO      : REAL := 2.0;       // 段中心除数 [-] / Zone centre divisor [-]
    DL_HALF     : REAL := 0.5;       // 插值区间归一化中点 [-] / Interpolation midpoint [-]
    DL_T_LO_C   : REAL := 0.0;       // 温度量程下限 [°C] / Temperature range low [°C]
    DL_T_HI_C   : REAL := 1200.0;    // 温度量程上限 [°C] / Temperature range high [°C]
    DL_ZONE_MAX : INT  := 1000;      // 段号钳制上限（防组态异常）[-] / Zone index ceiling [-]
END_VAR

(* —— 段 1：非有限值闸（R19：五路实值入参全覆盖，拦 NaN 与 Inf） —— *)
IF NOT (fT1C > -DL_BIG AND fT1C < DL_BIG)
   OR NOT (fT2C > -DL_BIG AND fT2C < DL_BIG)
   OR NOT (fT3C > -DL_BIG AND fT3C < DL_BIG)
   OR NOT (fZoneLenM > -DL_BIG AND fZoneLenM < DL_BIG)
   OR NOT (fZoneSpanM > -DL_BIG AND fZoneSpanM < DL_BIG) THEN
    fLocalC := 0.0;                         // 输出强制 0.0 / Output forced to zero
    fGradCpm := 0.0;                        // 梯度强制 0.0 / Gradient forced to zero
    iZoneClamp := 1;                        // 段号退到 1 / Zone index falls back to 1
    xValid := FALSE;                        // 有效位清零 / Validity cleared
    FC_DL_FloatBathTempProfileCalc := FALSE;   // 返回码同源 / Return mirrors validity
    RETURN;                                 // 立即退出 / Immediate exit
END_IF

(* —— 段 2：分母零闸（R4：总长与段长都是插值基准） —— *)
IF (ABS(fZoneLenM) <= DL_EPS) OR (ABS(fZoneSpanM) <= DL_EPS) THEN
    fLocalC := 0.0;                         // 输出强制 0.0 / Output forced to zero
    fGradCpm := 0.0;                        // 梯度强制 0.0 / Gradient forced to zero
    iZoneClamp := 1;                        // 段号退到 1 / Zone index falls back to 1
    xValid := FALSE;                        // 判无效 / Invalid
    FC_DL_FloatBathTempProfileCalc := FALSE;   // 返回码同步 / Return synchronised
    RETURN;                                 // 提前退出 / Early exit
END_IF

(* —— 段 3：负值闸（长度不可为负） —— *)
IF (fZoneLenM < 0.0) OR (fZoneSpanM < 0.0) THEN
    fLocalC := 0.0;                         // 输出强制 0.0 / Output forced to zero
    fGradCpm := 0.0;                        // 梯度强制 0.0 / Gradient forced to zero
    iZoneClamp := 1;                        // 段号退到 1 / Zone index falls back to 1
    xValid := FALSE;                        // 判无效 / Invalid
    FC_DL_FloatBathTempProfileCalc := FALSE;   // 返回码同步 / Return synchronised
    RETURN;                                 // 提前退出 / Early exit
END_IF

(* —— 段 4：段号钳制（1 ~ N 闭区间，N 由总长/段长取整，至少 1 段） —— *)
_iZoneCount := REAL_TO_INT(fZoneLenM / fZoneSpanM);               // 总段数 [-]（向下取整）
_iZoneCount := MAX(1, MIN(_iZoneCount, DL_ZONE_MAX));             // 段数钳 1..1000
iZoneClamp := MAX(1, MIN(iZone, _iZoneCount));                    // 段号钳 1..N

(* —— 段 5：位置归一化（R22 方向自核：段中心位置从 0 起算，除总长得 0..1） —— *)
_fPosM := (INT_TO_REAL(iZoneClamp - 1) * fZoneSpanM) + (fZoneSpanM / DL_TWO);   // 段中心 [m]
_fU := LIMIT(0.0, _fPosM / fZoneLenM, 1.0);                       // 归一化位置 [-]

(* —— 段 6：温度量程钳制 —— *)
_fT1Clamp := LIMIT(DL_T_LO_C, fT1C, DL_T_HI_C);                   // 入口温度钳 [°C]
_fT2Clamp := LIMIT(DL_T_LO_C, fT2C, DL_T_HI_C);                   // 中段温度钳 [°C]
_fT3Clamp := LIMIT(DL_T_LO_C, fT3C, DL_T_HI_C);                   // 出口温度钳 [°C]

(* —— 段 7：三段折线插值与区间梯度（u <= 0.5 属前区间，否则属后区间） —— *)
_fSegLenM := fZoneLenM * DL_HALF;                                 // 单区间物理长度 [m]
IF _iZoneCount <= 1 THEN
    _fLocalRaw := _fT1Clamp;                                      // 单段退化：取入口温度
    _fGradRaw := 0.0;                                             // 单段无梯度
ELSIF _fU <= DL_HALF THEN
    _fLocalRaw := _fT1Clamp + (_fT2Clamp - _fT1Clamp) * (_fU / DL_HALF);         // 前区间插值 [°C]
    _fGradRaw := (_fT2Clamp - _fT1Clamp) / _fSegLenM;                            // 前区间梯度 [°C/m]
ELSE
    _fLocalRaw := _fT2Clamp + (_fT3Clamp - _fT2Clamp) * ((_fU - DL_HALF) / DL_HALF);   // 后区间插值
    _fGradRaw := (_fT3Clamp - _fT2Clamp) / _fSegLenM;                            // 后区间梯度 [°C/m]
END_IF

(* —— 段 8：输出单点写盘（饱和钳制） —— *)
fLocalC := LIMIT(DL_T_LO_C, _fLocalRaw, DL_T_HI_C);               // 段温度 [°C]
fGradCpm := LIMIT(-DL_BIG, _fGradRaw, DL_BIG);                    // 梯度 [°C/m]

(* —— 段 9：有效位单点聚合（三个温度给定点在量程内） —— *)
xValid := (fT1C >= DL_T_LO_C) AND (fT1C <= DL_T_HI_C)
          AND (fT2C >= DL_T_LO_C) AND (fT2C <= DL_T_HI_C)
          AND (fT3C >= DL_T_LO_C) AND (fT3C <= DL_T_HI_C);
FC_DL_FloatBathTempProfileCalc := xValid;                         // 返回码：TRUE = 计算可信

END_FUNCTION

(* ---- FC_DL_FlocDilutionRatio.st ---- *)
(*
  道莅工业代码库 / Daoli Industrial ST Library
  组件: FC_DL_FlocDilutionRatio
  分类: DL_Process
  开源溯源: 无（clean-room 工程公式自研；参考公开工艺计算公式，未复制任何受版权保护代码）
  许可证: 本项目自有 (MIT)
  功能: 絮凝剂由高浓度母液稀释到目标浓度的稀释比与所需母液体积
*)
FUNCTION FC_DL_FlocDilutionRatio : BOOL
VAR_INPUT
    rStockPct : REAL; // 母液质量浓度 [%] / stock solution mass concentration
    rTargetPct : REAL; // 目标使用质量浓度 [%] / target working concentration
    rTankVolL : REAL; // 配液罐有效容积 [L] / dilution tank working volume
END_VAR
VAR_OUTPUT
    rRatio : REAL; // 稀释比 = 目标浓度/母液浓度 [L母液/L配液] / dilution ratio, stock litres per litre of batch
    rStockVolL : REAL; // 需投母液体积 [L] / required stock volume
    bValid : BOOL; // 结果有效位 [-] / result valid flag
    iErrCode : INT; // 事件码 0=正常 1=母液浓度非法 2=目标浓度高于母液已按 1:1 饱和 3=结果非有限 / event code
END_VAR
VAR
    rRatioUse : REAL; // 实际使用稀释比（含饱和修正）[L/L] / dilution ratio actually applied
END_VAR

    // —— 段 0：全路径预清 —— //
    rRatioUse := 0.0;
    rRatio := 0.0;
    rStockVolL := 0.0;
    bValid := FALSE;
    iErrCode := 0;
    FC_DL_FlocDilutionRatio := FALSE;
    // —— 段 1：分母闸（母液浓度） —— //
    IF ABS(rStockPct) <= 1.0E-9 THEN
        iErrCode := 1; // 母液浓度非法，稀释比无定义 / bad stock concentration, ratio undefined
        RETURN;
    END_IF;
    // —— 段 2：量纲链 (%),(%) 同量纲相除得无量纲比 [L母液/L配液] —— //
    rRatioUse := rTargetPct / rStockPct; // 稀释比 [-] / raw dilution ratio
    // —— 段 3：目标浓度不得高于母液（无法靠稀释提浓），按 1:1 饱和 —— //
    IF rTargetPct > rStockPct THEN
        rRatioUse := 1.0; // 饱和为纯母液 / saturate to neat stock
        iErrCode := 2; // 信息级：目标浓度超母液，已按 1:1 处理 / info: target above stock, clamped to 1:1
    END_IF;
    IF rRatioUse < 0.0 THEN
        rRatioUse := 0.0; // 负浓度输入防御 / negative concentration guard
    END_IF;
    rRatio := rRatioUse;
    // —— 段 4：配液体积换算与结果域闸 —— //
    rStockVolL := rTankVolL * rRatio; // 需母液体积 [L] / required stock volume
    IF (ABS(rStockVolL) > 1.0E15) OR (ABS(rRatio) > 1.0E15) THEN
        rStockVolL := 0.0;
        rRatio := 0.0;
        iErrCode := 3; // 结果非有限，强制归零 / non-finite result, forced to zero
        RETURN;
    END_IF;
    bValid := TRUE;
    FC_DL_FlocDilutionRatio := TRUE;
END_FUNCTION

(* ---- FC_DL_FoamSuppressDutyCalc.st ---- *)
(*
  ============================================================
  组件名 : FC_DL_FoamSuppressDutyCalc
  分类   : DL_Process
  功能   : 抑泡剂投加占空比计算，按液位抬高、灌装速率与基准投加量合成占空比并限幅
  复杂度 : C1
  版本   : 1.0.0
  作者   : 道莅工业代码库工厂 / R81
  日期   : 2026-11-24
  开源溯源 : clean-room（no upstream）—— 依据公开工程公式自研，未复制任何上游实现
  红线自检 : R1 无GVL/R2 无物理地址/R3 纯IEC/R4 防除零/R5 双语注释
  接口说明 :
      占空比 = 基准投加量 * (1 + 液位/100) * 灌装速率 / 100，结果限幅到 0~100。
      液位越高泡沫越易生成，故以液位对基准投加量做上浮修正；限幅保证输出可直接驱动 PWM。
  ============================================================
*)
FUNCTION FC_DL_FoamSuppressDutyCalc : BOOL
VAR_INPUT
    bEnable    : BOOL; // 使能：TRUE 时计算 / Enable: TRUE to compute
    bErr       : BOOL; // 外部故障：TRUE 时立即退出并置结果无效 / External fault: TRUE aborts with invalid result
    rLevelPct  : REAL; // 当前液位百分比 [%] / current liquid level [percent]
    rFillRate  : REAL; // 灌装体积速率 [L/min] / filling volumetric rate [litre per minute]
    rDoseBase  : REAL; // 基准投加量 [mL/L] / base dosing quantity [millilitre per litre]
END_VAR
VAR_OUTPUT
    rDutyPct     : REAL; // 抑泡投加占空比，限幅 0~100 [%] / foam suppression duty cycle clamped to 0 to 100 [percent]
    rDoseRawPct  : REAL; // 限幅前的原始占空比 [%] / raw duty cycle before clamping [percent]
    bClamped     : BOOL; // 限幅生效：TRUE 表示输出被截断 / clamping active, TRUE means the output was truncated
    bValid       : BOOL; // 输出有效：TRUE 表示结果可用 / Output valid
END_VAR
VAR CONSTANT
    DL_R_MAX  : REAL := 3.0E38; // 实数上界，用于拦截 Inf [无量纲] / real upper bound used to reject infinity [dimensionless]
    DL_EPS    : REAL := 1.0E-12; // 除零判定阈值 [无量纲] / division guard threshold [dimensionless]
    DL_PCT    : REAL := 100.0;   // 百分数换算系数 [无量纲] / percentage scaling factor [dimensionless]
    DL_DUTY_HI : REAL := 100.0;  // 占空比上限 [%] / duty cycle upper limit [percent]
    DL_DUTY_LO : REAL := 0.0;    // 占空比下限 [%] / duty cycle lower limit [percent]
    DL_LEVEL_HI : REAL := 100.0; // 液位允许上限 [%] / permitted upper bound of the level [percent]
END_VAR
VAR
    _bFin : BOOL := FALSE; // 输入有限性判定结果 / input finiteness verdict
    _rLvl : REAL := 0.0;   // 液位修正系数 [无量纲] / level correction factor [dimensionless]
END_VAR

    // 段 1｜出口预置
    rDutyPct := 0.0;
    rDoseRawPct := 0.0;
    bClamped := FALSE;
    bValid := FALSE;
    // 段 2｜使能闸与外部故障闸
    IF NOT bEnable THEN
        RETURN;
    END_IF;
    IF bErr THEN
        RETURN;
    END_IF;
    // 段 3｜非有限闸
    _bFin := (rLevelPct = rLevelPct) AND (ABS(rLevelPct) <= DL_R_MAX) AND (rFillRate = rFillRate) AND (ABS(rFillRate) <= DL_R_MAX) AND (rDoseBase = rDoseBase) AND (ABS(rDoseBase) <= DL_R_MAX);
    IF NOT _bFin THEN
        RETURN;
    END_IF;
    // 段 4｜域闸：液位 0~100，速率与投加量不得为负
    IF (rLevelPct < DL_DUTY_LO) OR (rLevelPct > DL_LEVEL_HI) THEN
        RETURN;
    END_IF;
    IF (rFillRate < DL_DUTY_LO) OR (rDoseBase < DL_DUTY_LO) THEN
        RETURN;
    END_IF;
    // 段 5｜主体合成：液位越高修正系数越大
    _rLvl := 1.0 + rLevelPct / DL_PCT;
    rDoseRawPct := rDoseBase * _rLvl * rFillRate / DL_PCT;
    // 段 6｜限幅并记录截断标志
    IF rDoseRawPct > DL_DUTY_HI THEN
        rDutyPct := DL_DUTY_HI;
        bClamped := TRUE;
    ELSIF rDoseRawPct < DL_DUTY_LO THEN
        rDutyPct := DL_DUTY_LO;
        bClamped := TRUE;
    ELSE
        rDutyPct := rDoseRawPct;
        bClamped := FALSE;
    END_IF;
    bValid := TRUE;
    FC_DL_FoamSuppressDutyCalc := bValid;
END_FUNCTION

(* ---- FC_DL_ForgeBilletHeatTimeCalc.st ---- *)
(*
  Name: FC_DL_ForgeBilletHeatTimeCalc
  Category: DL_Process
  Version: 1.0.0
  Round: R89 / 2026-11-25
  开源溯源：clean-room 自研（族 锻造加热退火，ST 开源生态实测 0 命中，无外部代码引入）
  功能：坯料加热时间（透热厚度经验式）：以加热系数乘透热厚度，并按炉温-目标温差势比修正，另给出均热时间。
  边界条件：① 五入参全部过非有限闸，任一非有限返回哨兵 -1；
            ② 炉温必须高于目标温度（否则无传热势差，返回哨兵 -1），目标温度必须高于起始温度；
            ③ 势比 = (T炉−T初)/(T炉−T目标)：目标温度越接近炉温，势比越大（加热越慢），量纲无量纲；
            ④ 均热时间取加热时间的 25 %，并设 5 min 下限（薄料均热不因比例过小而失效）。
  量纲自证：k[min/cm] × 厚度[cm] = min；势比无量纲，量纲保持 min。
*)
FUNCTION FC_DL_ForgeBilletHeatTimeCalc : REAL
VAR_INPUT
    fThkMm : REAL;              (* 坯料透热厚度 [mm] Billet through-heating thickness [mm] *)
    fHeatCoefMinPerCm : REAL;   (* 加热系数 [min/cm] Heating coefficient [min/cm] *)
    fFurnaceTempC : REAL;       (* 炉膛温度 [℃] Furnace temperature [degC] *)
    fTargetTempC : REAL;        (* 目标出炉温度 [℃] Target discharge temperature [degC] *)
    fStartTempC : REAL;         (* 入炉起始温度 [℃] Charging temperature [degC] *)
END_VAR
VAR_OUTPUT
    fHeatTimeMin : REAL;        (* 加热时间 [min] Heating time [min] *)
    fSoakTimeMin : REAL;        (* 均热时间 [min] Soak time [min] *)
    xValid : BOOL;              (* 计算有效性标志 [-] Calculation valid flag *)
END_VAR
VAR CONSTANT
    DL_EPS : REAL := 1.0E-9;        (* 判据容差 [-] Criterion tolerance *)
    DL_MM_PER_CM : REAL := 10.0;    (* 毫米 → 厘米换算 [mm/cm] Millimetre to centimetre *)
    DL_SOAK_RATIO : REAL := 0.25;   (* 均热/加热时间比 [-] Soak to heat ratio *)
    DL_SOAK_MIN : REAL := 5.0;      (* 均热时间下限 [min] Soak time floor [min] *)
    DL_T_MIN : REAL := 10.0;        (* 厚度下限 [mm] Thickness floor [mm] *)
    DL_T_MAX : REAL := 1200.0;      (* 厚度上限 [mm] Thickness ceiling [mm] *)
    DL_K_MIN : REAL := 0.5;         (* 加热系数下限 [min/cm] Coefficient floor [min/cm] *)
    DL_K_MAX : REAL := 10.0;        (* 加热系数上限 [min/cm] Coefficient ceiling [min/cm] *)
    DL_F_MIN : REAL := 200.0;       (* 炉温下限 [℃] Furnace floor [degC] *)
    DL_F_MAX : REAL := 1400.0;      (* 炉温上限 [℃] Furnace ceiling [degC] *)
    DL_S_MIN : REAL := -50.0;       (* 起始温度下限 [℃] Start floor [degC] *)
    DL_S_MAX : REAL := 1200.0;      (* 起始温度上限 [℃] Start ceiling [degC] *)
END_VAR
VAR
    fThkCm : REAL;      (* 透热厚度 [cm] Through-heating thickness [cm] *)
    fPotRatio : REAL;   (* 温差势比 [-] Temperature potential ratio *)
    fDenC : REAL;       (* 势比分母（炉温−目标） [℃] Potential denominator [degC] *)
END_VAR
(* 出口预置：三出口统一预置（R256） *)
fHeatTimeMin := 0.0; fSoakTimeMin := 0.0; xValid := FALSE;
(* 非有限闸：NaN 自反判 + Inf 差值自减判，五入参全枚举 *)
IF (fThkMm <> fThkMm) OR ((fThkMm - fThkMm) <> 0.0)
   OR (fHeatCoefMinPerCm <> fHeatCoefMinPerCm) OR ((fHeatCoefMinPerCm - fHeatCoefMinPerCm) <> 0.0)
   OR (fFurnaceTempC <> fFurnaceTempC) OR ((fFurnaceTempC - fFurnaceTempC) <> 0.0)
   OR (fTargetTempC <> fTargetTempC) OR ((fTargetTempC - fTargetTempC) <> 0.0)
   OR (fStartTempC <> fStartTempC) OR ((fStartTempC - fStartTempC) <> 0.0) THEN
    FC_DL_ForgeBilletHeatTimeCalc := -1.0;  (* 哨兵 -1：入参非有限 / Sentinel -1, non-finite input *)
    RETURN;
END_IF
(* 组态域闸：厚度、系数、炉温、起始温度定域，温度须满足 炉温 > 目标 > 起始 *)
IF (fThkMm < DL_T_MIN) OR (fThkMm > DL_T_MAX)
   OR (fHeatCoefMinPerCm < DL_K_MIN) OR (fHeatCoefMinPerCm > DL_K_MAX)
   OR (fFurnaceTempC < DL_F_MIN) OR (fFurnaceTempC > DL_F_MAX)
   OR (fStartTempC < DL_S_MIN) OR (fStartTempC > DL_S_MAX)
   OR (fTargetTempC <= fStartTempC) OR ((fFurnaceTempC - fTargetTempC) <= DL_EPS) THEN
    FC_DL_ForgeBilletHeatTimeCalc := -1.0;  (* 哨兵 -1：组态非法 / Sentinel -1, bad configuration *)
    RETURN;
END_IF
(* 透热厚度折算：mm ÷ 10 = cm *)
fThkCm := fThkMm / DL_MM_PER_CM;
(* 势比：分母（炉温−目标）已过正性闸，绝无零除 *)
fDenC := fFurnaceTempC - fTargetTempC;
fPotRatio := (fFurnaceTempC - fStartTempC) / fDenC;
(* 加热时间：k[min/cm] × 厚度[cm] × 势比，量纲 min *)
fHeatTimeMin := fHeatCoefMinPerCm * fThkCm * fPotRatio;
(* 均热时间：25 % 加热时间，并保 5 min 下限 *)
fSoakTimeMin := fHeatTimeMin * DL_SOAK_RATIO;
IF fSoakTimeMin < DL_SOAK_MIN THEN
    fSoakTimeMin := DL_SOAK_MIN;            (* 下限钳位 / Floor clamp *)
END_IF
xValid := TRUE;                             (* 链路有效 / Chain valid *)
FC_DL_ForgeBilletHeatTimeCalc := fHeatTimeMin;
END_FUNCTION

(* ---- FC_DL_ForgeLoadTonCalc.st ---- *)
(*
  Name: FC_DL_ForgeLoadTonCalc
  Category: DL_Process
  Version: 1.0.0
  Round: R89 / 2026-11-25
  开源溯源：clean-room 自研（族 锻造加热退火，ST 开源生态实测 0 命中，无外部代码引入）
  功能：锻造载荷：投影面积 × 变形抗力 × 形状系数得锻造力，折算吨位与压机利用率。
  边界条件：① 三入参全部过非有限闸，任一非有限返回哨兵 -1；
            ② 投影面积 100~5e6 mm2、变形抗力 20~400 MPa、形状系数 1.0~3.0 为工程域，越域返回哨兵 -1；
            ③ 压机额定载荷为常量 DL_FLT_PRESS_KN（默认 20000 kN），利用率可超 100 %（超载照实上报不钳位）。
  量纲自证：mm2 × (N/mm2) = N；N/1000 = kN；kN ÷ 9.80665[kN/tf] = tf 折算吨位。
*)
FUNCTION FC_DL_ForgeLoadTonCalc : REAL
VAR_INPUT
    fProjAreaMm2 : REAL;        (* 锻件投影面积 [mm2] Forging projected area [mm2] *)
    fFlowStressMpa : REAL;      (* 变形抗力（流动应力） [MPa] Flow stress [MPa] *)
    fShapeFactor : REAL;        (* 形状系数（1.0~3.0） [-] Shape factor *)
END_VAR
VAR_OUTPUT
    fLoadKN : REAL;             (* 锻造力 [kN] Forging load [kN] *)
    fLoadTon : REAL;            (* 折算吨位 [tf] Load in tonne-force [tf] *)
    fPressUtilPct : REAL;       (* 压机利用率（可超 100 %） [%] Press utilization [%] *)
    xValid : BOOL;              (* 计算有效性标志 [-] Calculation valid flag *)
END_VAR
VAR CONSTANT
    DL_KN_PER_N : REAL := 1000.0;       (* 牛 → 千牛换算 [N/kN] Newton to kilonewton *)
    DL_KN_PER_TF : REAL := 9.80665;     (* 吨力 → 千牛换算 [kN/tf] Kilonewton per tonne-force *)
    DL_FLT_PRESS_KN : REAL := 20000.0;  (* 压机额定载荷（可改常量） [kN] Press rated load [kN] *)
    DL_PCT : REAL := 100.0;             (* 百分数基准 [%] Percent base *)
    DL_A_MIN : REAL := 100.0;           (* 投影面积下限 [mm2] Area floor [mm2] *)
    DL_A_MAX : REAL := 5000000.0;       (* 投影面积上限 [mm2] Area ceiling [mm2] *)
    DL_S_MIN : REAL := 20.0;            (* 变形抗力下限 [MPa] Flow stress floor [MPa] *)
    DL_S_MAX : REAL := 400.0;           (* 变形抗力上限 [MPa] Flow stress ceiling [MPa] *)
    DL_F_MIN : REAL := 1.0;             (* 形状系数下限 [-] Shape factor floor *)
    DL_F_MAX : REAL := 3.0;             (* 形状系数上限 [-] Shape factor ceiling *)
END_VAR
VAR
    fForceN : REAL;     (* 锻造力（牛） [N] Forging force [N] *)
END_VAR
(* 出口预置：四出口统一预置（R256） *)
fLoadKN := 0.0; fLoadTon := 0.0; fPressUtilPct := 0.0; xValid := FALSE;
(* 非有限闸：NaN 自反判 + Inf 差值自减判，三入参全枚举 *)
IF (fProjAreaMm2 <> fProjAreaMm2) OR ((fProjAreaMm2 - fProjAreaMm2) <> 0.0)
   OR (fFlowStressMpa <> fFlowStressMpa) OR ((fFlowStressMpa - fFlowStressMpa) <> 0.0)
   OR (fShapeFactor <> fShapeFactor) OR ((fShapeFactor - fShapeFactor) <> 0.0) THEN
    FC_DL_ForgeLoadTonCalc := -1.0;         (* 哨兵 -1：入参非有限 / Sentinel -1, non-finite input *)
    RETURN;
END_IF
(* 组态域闸：面积、变形抗力、形状系数逐项定域 *)
IF (fProjAreaMm2 < DL_A_MIN) OR (fProjAreaMm2 > DL_A_MAX)
   OR (fFlowStressMpa < DL_S_MIN) OR (fFlowStressMpa > DL_S_MAX)
   OR (fShapeFactor < DL_F_MIN) OR (fShapeFactor > DL_F_MAX) THEN
    FC_DL_ForgeLoadTonCalc := -1.0;         (* 哨兵 -1：组态非法 / Sentinel -1, bad configuration *)
    RETURN;
END_IF
(* 锻造力：mm2 × N/mm2 = N，再乘无量纲形状系数 *)
fForceN := fProjAreaMm2 * fFlowStressMpa * fShapeFactor;
(* 折算 kN 与吨位：kN ÷ kN/tf = tf *)
fLoadKN := fForceN / DL_KN_PER_N;
fLoadTon := fLoadKN / DL_KN_PER_TF;
(* 压机利用率：常量额定载荷恒正，超载照实超 100 %（事实不钳位） *)
fPressUtilPct := (fLoadKN / DL_FLT_PRESS_KN) * DL_PCT;
xValid := TRUE;                             (* 链路有效 / Chain valid *)
FC_DL_ForgeLoadTonCalc := fLoadKN;
END_FUNCTION

(* ---- FC_DL_ForkExtendSafeChk.st ---- *)
(*
  ============================================================
  组件名 : FC_DL_ForkExtendSafeChk
  分类   : DL_Process
  功能   : 货叉伸出安全校核，同时校验通道余量是否足够与货位对齐误差是否在容差内
  复杂度 : C1
  版本   : 1.0.0
  作者   : 道莅工业代码库工厂 / R81
  日期   : 2026-11-24
  开源溯源 : clean-room（no upstream）—— 依据公开工程公式自研，未复制任何上游实现
  红线自检 : R1 无GVL/R2 无物理地址/R3 纯IEC/R4 防除零/R5 双语注释
  接口说明 :
      安全判据必须两条同时满足：需伸量 <= 通道余量 - 安全余量，且对齐误差绝对值 <= 容差。
      余量 rMargin_mm = 通道余量 - 安全余量 - 需伸量，为负表示越界，正值表示剩余空间。
      任一条不满足即 bSafe=FALSE，同时 bValid 仍为 TRUE，因为判定结论本身是确定的。
  ============================================================
*)
FUNCTION FC_DL_ForkExtendSafeChk : BOOL
VAR_INPUT
    bEnable        : BOOL; // 使能：TRUE 时校核 / Enable: TRUE to check
    bErr           : BOOL; // 外部故障：TRUE 时立即退出并置结果无效 / External fault: TRUE aborts with invalid result
    rForkExt_mm    : REAL; // 本次需要伸出的货叉长度 [mm] / required fork extension for this cycle [mm]
    rAisleClear_mm : REAL; // 巷道侧向可用余量 [mm] / available lateral clearance in the aisle [mm]
    rAlignErr_mm   : REAL; // 货位对齐误差，带正负号 [mm] / cell alignment error with sign [mm]
    rAlignTol_mm   : REAL; // 允许的对齐误差容差 [mm] / permitted alignment tolerance [mm]
    rSafeMargin_mm : REAL; // 需保留的安全余量 [mm] / safety margin that must be preserved [mm]
END_VAR
VAR_OUTPUT
    bSafe      : BOOL; // 伸出安全：TRUE 表示两条判据同时满足 / extension safe, TRUE when both criteria hold
    rMargin_mm : REAL; // 伸出后剩余余量，负值表示越界 [mm] / remaining margin after extension, negative means overrun [mm]
    bAlignOk   : BOOL; // 对齐合格：TRUE 表示误差在容差内 / alignment acceptable, TRUE when the error is within tolerance
    bValid     : BOOL; // 输出有效：TRUE 表示结果可用 / Output valid
END_VAR
VAR CONSTANT
    DL_R_MAX : REAL := 3.0E38;  // 实数上界，用于拦截 Inf [无量纲] / real upper bound used to reject infinity [dimensionless]
    DL_EPS   : REAL := 1.0E-12; // 除零判定阈值 [无量纲] / division guard threshold [dimensionless]
    DL_ZERO  : REAL := 0.0;     // 零值常量 [无量纲] / zero constant [dimensionless]
END_VAR
VAR
    _bFin    : BOOL := FALSE; // 输入有限性判定结果 / input finiteness verdict
    _rAllow  : REAL := 0.0;   // 扣掉安全余量后的可伸长度 [mm] / allowable extension after removing the safety margin [mm]
    _rAbsErr : REAL := 0.0;   // 对齐误差绝对值 [mm] / absolute alignment error [mm]
END_VAR

    // 段 1｜出口预置：安全位保守置 FALSE，余量置零
    bSafe := FALSE;
    rMargin_mm := 0.0;
    bAlignOk := FALSE;
    bValid := FALSE;
    // 段 2｜使能闸与外部故障闸
    IF NOT bEnable THEN
        RETURN;
    END_IF;
    IF bErr THEN
        RETURN;
    END_IF;
    // 段 3｜非有限闸
    _bFin := (rForkExt_mm = rForkExt_mm) AND (ABS(rForkExt_mm) <= DL_R_MAX) AND (rAisleClear_mm = rAisleClear_mm) AND (ABS(rAisleClear_mm) <= DL_R_MAX) AND (rAlignErr_mm = rAlignErr_mm) AND (ABS(rAlignErr_mm) <= DL_R_MAX) AND (rAlignTol_mm = rAlignTol_mm) AND (ABS(rAlignTol_mm) <= DL_R_MAX) AND (rSafeMargin_mm = rSafeMargin_mm) AND (ABS(rSafeMargin_mm) <= DL_R_MAX);
    IF NOT _bFin THEN
        RETURN;
    END_IF;
    // 段 4｜域闸：需伸量、通道余量、容差、安全余量均不得为负
    IF (rForkExt_mm < DL_ZERO) OR (rAisleClear_mm < DL_ZERO) OR (rAlignTol_mm < DL_ZERO) OR (rSafeMargin_mm < DL_ZERO) THEN
        RETURN;
    END_IF;
    // 段 5｜可伸长度与剩余余量
    _rAllow := rAisleClear_mm - rSafeMargin_mm;
    rMargin_mm := _rAllow - rForkExt_mm;
    // 段 6｜两条判据
    _rAbsErr := ABS(rAlignErr_mm);
    IF _rAbsErr <= rAlignTol_mm THEN
        bAlignOk := TRUE;
    ELSE
        bAlignOk := FALSE;
    END_IF;
    IF (rForkExt_mm <= _rAllow) AND bAlignOk THEN
        bSafe := TRUE;
    ELSE
        bSafe := FALSE;
    END_IF;
    bValid := TRUE;
    FC_DL_ForkExtendSafeChk := bValid;
END_FUNCTION

(* ---- FC_DL_GasHolderLevel.st ---- *)
(*
  道莅工业代码库 / Daoli Industrial ST Library
  组件: FC_DL_GasHolderLevel
  分类: DL_Process
  开源溯源: 无（clean-room 工程公式自研；参考公开工艺计算公式，未复制任何受版权保护代码）
  许可证: 本项目自有 (MIT)
  功能: 湿式气柜储气量标态折算与可释放能量估算
  口径声明: 能量按厂内标定简化系数 0.55 kWh/(m3·单位甲烷份额)×CH4 假设 0.6 计，
            非热力学严格值（严格口径为 9.94 kWh/m3 纯甲烷），仅供储量看板同比使用
*)
FUNCTION FC_DL_GasHolderLevel : BOOL
VAR_INPUT
    rPressKpa : REAL; // 柜内表压 [kPa] / gauge pressure in the holder
    rTempC : REAL; // 柜内气体温度 [°C] / gas temperature
    rVolM3 : REAL; // 气柜几何容积 [m3] / geometric holder volume
    rLevelPct : REAL; // 有效储气液位/行程 [%] / effective storage level
END_VAR
VAR_OUTPUT
    rNormM3 : REAL; // 标态储气量 [Nm3] / normalised stored volume
    rEnergyKwh : REAL; // 可释放能量估算 [kWh] / estimated releasable energy
    bValid : BOOL; // 结果有效位 [-] / result valid flag
    iErrCode : INT; // 事件码 0=正常 1=温度超域 2=容积非法 3=压力非法 4=结果非有限 / event code
END_VAR
VAR CONSTANT
    rKelvinOff : REAL := 273.15; // 开尔文偏移 [K] / kelvin offset
    rPressRefKpa : REAL := 101.325; // 标准大气压 [kPa] / standard atmospheric pressure
    rTempMinC : REAL := -50.0; // 温度域下限 [°C] / temperature lower bound
    rPctToFrac : REAL := 0.01; // 百分数转小数系数 [-]/[%] / percent to fraction factor
    rKwhPerM3 : REAL := 0.55; // 能量简化系数 [kWh/m3] / simplified energy coefficient
    rCh4Assumed : REAL := 0.6; // 甲烷份额假设 [-] / assumed methane fraction
END_VAR
VAR
    rTempK : REAL; // 柜内绝对温度 [K] / absolute temperature
    rVolUseM3 : REAL; // 有效储气体积 [m3] / effective stored volume
    rNormRaw : REAL; // 未校验标态量 [Nm3] / unchecked normalised volume
END_VAR

    // —— 段 0：全路径预清 —— //
    rTempK := 0.0;
    rVolUseM3 := 0.0;
    rNormRaw := 0.0;
    rNormM3 := 0.0;
    rEnergyKwh := 0.0;
    bValid := FALSE;
    iErrCode := 0;
    FC_DL_GasHolderLevel := FALSE;
    // —— 段 1：温度域闸（同时保护标态折算分母 273.15+T） —— //
    IF rTempC <= rTempMinC THEN
        iErrCode := 1; // 温度超域，标态折算无意义 / temperature out of domain
        RETURN;
    END_IF;
    IF rVolM3 <= 0.0 THEN
        iErrCode := 2; // 容积非法 / invalid holder volume
        RETURN;
    END_IF;
    // —— 段 2：压力域闸（表压需为正，绝对压 = 表压 + 大气压） —— //
    IF rPressKpa <= 0.0 THEN
        iErrCode := 3; // 压力非法，绝对压不可信 / invalid gauge pressure
        RETURN;
    END_IF;
    // —— 段 3：有效储气体积按液位折算，再作标态换算（量纲 m3×kPa/K÷kPa = Nm3） —— //
    rVolUseM3 := rVolM3 * rLevelPct * rPctToFrac; // 有效体积 [m3] / effective volume
    IF rVolUseM3 < 0.0 THEN
        rVolUseM3 := 0.0; // 负液位防御 / negative level guard
    END_IF;
    rTempK := rKelvinOff + rTempC; // 绝对温度 [K] / absolute temperature
    rNormRaw := rVolUseM3 * (rPressRefKpa + rPressKpa) * rKelvinOff / (rTempK * rPressRefKpa); // 标态量 [Nm3]
    IF ABS(rNormRaw) > 1.0E15 THEN
        iErrCode := 4; // 结果非有限，强制归零 / non-finite result, forced to zero
        RETURN;
    END_IF;
    rNormM3 := rNormRaw;
    // —— 段 4：能量估算（量纲 Nm3 × kWh/m3 × - = kWh） —— //
    rEnergyKwh := rNormM3 * rKwhPerM3 * rCh4Assumed; // 能量估算 [kWh] / estimated energy
    bValid := TRUE;
    FC_DL_GasHolderLevel := TRUE;
END_FUNCTION

(* ---- FC_DL_GlassCutOptimizeCalc.st ---- *)
(*
  Name: FC_DL_GlassCutOptimizeCalc
  Category: DL_Process
  Version: 1.0.0
  Round: R90 / 2026-11-25
  开源溯源：clean-room 自研（族 浮法玻璃锡槽退火，ST 开源生态实测 0 命中，无外部代码引入）
  功能：1) 两种订单长度的最优切裁组合求解。枚举法而非贪心：把 A 规格的切裁数量从 0 穷举到
           订单需求上限，对每个 A 数量在剩余原板长度内按整除算出 B 规格的最大可切数量
           （再受 B 订单需求上限约束），得到该组合的实际用料长度；取全部组合中用料最长者。
           对两种规格的原板一维下料问题，穷举 A 数量 + 每档取最大 B 即为严格最优
           （每档内 B 取最大不会减少用料，且全部 A 档位已覆盖）。
        2) 余料率与利用率：利用率 fUtilPct = 最优用料 / 原板长度 × 100，
           余料 fScrapM = 原板长度 − 最优用料。余料必然 >= 0（穷举解保证不超原板）。
        3) 循环上界由订单需求与 DL_MAX_CNT 双重钳制，避免运行时无界循环拖垮扫描周期。
  边界条件：1) 非有限值闸：五个实值入参统一过 NOT(x > -DL_BIG AND x < DL_BIG)，
           同时拦 NaN 与 Inf，命中即拦断实值通路（两个 REAL 输出强制 0.0）并置无效（R19）。
        2) 分母零闸：原板长度与两种订单长度都必须 ABS > DL_EPS（任为 0 则整除与利用率无定义）。
        3) 负值闸：原板长度、两种订单长度为负，或两种数量为负均判无效
           （负数量无物理意义，取绝对值会虚增切裁方案）。
        4) 钳制：订单数量先钳到 0 ~ DL_MAX_CNT(200)，原板长度钳 0 ~ DL_LEN_MAX(100000 m)；
           数量被钳或原板越域时置 xValid=FALSE，避免把截断后的方案当作真实方案下发。
        5) 循环规范（R18）：只使用 FOR i := a TO b DO 的递增形式，禁用 DOWNTO。
  量纲自证：用料 = 段 × m + 段 × m = m；余料 = m − m = m；
           利用率 = m / m × 100 = 无因次 [%]，分子分母同量纲；
           整除式 _fRemain / fOrderLenB 得「段数」（无因次个数），再取整后乘回长度得 m。
*)

FUNCTION FC_DL_GlassCutOptimizeCalc : BOOL
VAR_INPUT
    fRibbonLenM   : REAL;   // 原板（玻璃带）可用长度 [m] / Available ribbon length [m]
    fOrderLenA    : REAL;   // A 规格订单长度 [m] / Order length A [m]
    fOrderLenB    : REAL;   // B 规格订单长度 [m] / Order length B [m]
    iQtyA         : INT;    // A 规格需求数量 [段] / Order quantity A [pcs]
    iQtyB         : INT;    // B 规格需求数量 [段] / Order quantity B [pcs]
END_VAR
VAR_OUTPUT
    fUtilPct      : REAL;   // 最优利用率 [%] / Optimal utilization ratio [%]
    fScrapM       : REAL;   // 余料长度 [m] / Scrap length [m]
    iBestA        : INT;    // 最优方案中的 A 数量 [段] / Quantity A in optimal plan [pcs]
    iBestB        : INT;    // 最优方案中的 B 数量 [段] / Quantity B in optimal plan [pcs]
    xValid        : BOOL;   // 计算有效标志 [bool] / Calculation valid flag [bool]
END_VAR
VAR
    _i                : INT;    // 枚举循环变量（A 规格数量）[段] / Enumeration index for A [pcs]
    _iQtyAClamp       : INT;    // 钳制后的 A 需求数量 [段] / Clamped quantity A [pcs]
    _iQtyBClamp       : INT;    // 钳制后的 B 需求数量 [段] / Clamped quantity B [pcs]
    _iBestACalc       : INT;    // 计算过程中的最优 A 数量 [段] / Best A during search [pcs]
    _iBestBCalc       : INT;    // 计算过程中的最优 B 数量 [段] / Best B during search [pcs]
    _iBMax            : INT;    // 当前 A 档位下 B 的可切数量 [段] / Max B at current A [pcs]
    _fRemainM         : REAL;   // 切完 A 后的剩余长度 [m] / Remaining length after A [m]
    _fUsedM           : REAL;   // 当前组合的实际用料 [m] / Used length of current plan [m]
    _fBestUsedM       : REAL;   // 已找到的最优用料 [m] / Best used length found [m]
    _fRibbonClamp     : REAL;   // 钳制后的原板长度 [m] / Clamped ribbon length [m]
    _fUtilRawPct      : REAL;   // 未饱和的利用率 [%] / Raw utilization ratio [%]
    _iQtyAMax         : INT;    // A 需求上限（钳制用）[段] / Quantity A ceiling [pcs]
    _iQtyBMax         : INT;    // B 需求上限（钳制用）[段] / Quantity B ceiling [pcs]
    _fQtyMaxReal      : REAL;   // 数量上限的实数形态 [段] / Quantity ceiling as real [pcs]
END_VAR
VAR CONSTANT
    DL_EPS        : REAL := 1.0E-9;    // 分母零闸阈值 [-] / Division-zero gate threshold [-]
    DL_BIG        : REAL := 1.0E12;    // 非有限值闸量级上限 [-] / Finiteness gate magnitude [-]
    DL_PCT        : REAL := 100.0;     // 百分比换算因子 [%] / Percent conversion factor [%]
    DL_MAX_CNT    : INT  := 200;       // 枚举与数量的钳制上限 [段] / Enumeration and quantity ceiling [pcs]
    DL_LEN_MAX    : REAL := 100000.0;  // 原板长度饱和上限 [m] / Ribbon length saturation ceiling [m]
END_VAR

(* —— 段 1：非有限值闸（R19：五路实值入参全覆盖，拦 NaN 与 Inf） —— *)
IF NOT (fRibbonLenM > -DL_BIG AND fRibbonLenM < DL_BIG)
   OR NOT (fOrderLenA > -DL_BIG AND fOrderLenA < DL_BIG)
   OR NOT (fOrderLenB > -DL_BIG AND fOrderLenB < DL_BIG) THEN
    fUtilPct := 0.0;                        // 输出强制 0.0 / Output forced to zero
    fScrapM := 0.0;                         // 余料强制 0.0 / Scrap forced to zero
    iBestA := 0;                            // 最优 A 数量清零 / Best A cleared
    iBestB := 0;                            // 最优 B 数量清零 / Best B cleared
    xValid := FALSE;                        // 有效位清零 / Validity cleared
    FC_DL_GlassCutOptimizeCalc := FALSE;    // 返回码同源 / Return mirrors validity
    RETURN;                                 // 立即退出 / Immediate exit
END_IF

(* —— 段 2：分母零闸（R4：原板长度与两种订单长度都是整除/归一的分母） —— *)
IF (ABS(fRibbonLenM) <= DL_EPS) OR (ABS(fOrderLenA) <= DL_EPS) OR (ABS(fOrderLenB) <= DL_EPS) THEN
    fUtilPct := 0.0;                        // 输出强制 0.0 / Output forced to zero
    fScrapM := 0.0;                         // 余料强制 0.0 / Scrap forced to zero
    iBestA := 0;                            // 最优 A 数量清零 / Best A cleared
    iBestB := 0;                            // 最优 B 数量清零 / Best B cleared
    xValid := FALSE;                        // 判无效 / Invalid
    FC_DL_GlassCutOptimizeCalc := FALSE;    // 返回码同步 / Return synchronised
    RETURN;                                 // 提前退出 / Early exit
END_IF

(* —— 段 3：负值闸（长度与数量均不可为负） —— *)
IF (fRibbonLenM < 0.0) OR (fOrderLenA < 0.0) OR (fOrderLenB < 0.0)
   OR (iQtyA < 0) OR (iQtyB < 0) THEN
    fUtilPct := 0.0;                        // 输出强制 0.0 / Output forced to zero
    fScrapM := 0.0;                         // 余料强制 0.0 / Scrap forced to zero
    iBestA := 0;                            // 最优 A 数量清零 / Best A cleared
    iBestB := 0;                            // 最优 B 数量清零 / Best B cleared
    xValid := FALSE;                        // 判无效 / Invalid
    FC_DL_GlassCutOptimizeCalc := FALSE;    // 返回码同步 / Return synchronised
    RETURN;                                 // 提前退出 / Early exit
END_IF

(* —— 段 4：数量与长度钳制（枚举上界必须是有界常量，禁止运行期无界循环） —— *)
_iQtyAMax := DL_MAX_CNT;                                          // A 需求上限 [段]
_iQtyBMax := DL_MAX_CNT;                                          // B 需求上限 [段]
_iQtyAClamp := MAX(0, MIN(iQtyA, _iQtyAMax));                     // 钳制后的 A 数量 [段]
_iQtyBClamp := MAX(0, MIN(iQtyB, _iQtyBMax));                     // 钳制后的 B 数量 [段]
_fRibbonClamp := LIMIT(0.0, fRibbonLenM, DL_LEN_MAX);             // 原板长度钳制 [m]
_fQtyMaxReal := INT_TO_REAL(DL_MAX_CNT);                          // 数量上限实数形态 [段]

(* —— 段 5：枚举最优切裁（R18：仅递增 FOR；A 档位穷举，每档 B 取最大） —— *)
_fBestUsedM := 0.0;                                               // 最优用料初值 [m]
_iBestACalc := 0;                                                 // 最优 A 初值 [段]
_iBestBCalc := 0;                                                 // 最优 B 初值 [段]
FOR _i := 0 TO _iQtyAClamp DO
    _fRemainM := _fRibbonClamp - INT_TO_REAL(_i) * fOrderLenA;    // 切 A 后的剩余长度 [m]
    IF _fRemainM >= 0.0 THEN
        _iBMax := REAL_TO_INT(LIMIT(0.0, _fRemainM / fOrderLenB, _fQtyMaxReal));   // B 可切数 [段]
        _iBMax := MIN(_iBMax, _iQtyBClamp);                       // 再受 B 需求上限约束
        _fUsedM := INT_TO_REAL(_i) * fOrderLenA + INT_TO_REAL(_iBMax) * fOrderLenB;   // 实际用料 [m]
        IF _fUsedM > _fBestUsedM THEN
            _fBestUsedM := _fUsedM;                               // 刷新最优用料
            _iBestACalc := _i;                                    // 记录最优 A 数量
            _iBestBCalc := _iBMax;                                // 记录最优 B 数量
        END_IF
    END_IF
END_FOR

(* —— 段 6：输出单点写盘（利用率与余料同源于 _fBestUsedM，保证两值自洽） —— *)
_fUtilRawPct := _fBestUsedM / _fRibbonClamp * DL_PCT;             // 利用率 [%]
fUtilPct := LIMIT(0.0, _fUtilRawPct, DL_PCT);                     // 利用率钳 0..100 [%]
fScrapM := LIMIT(0.0, _fRibbonClamp - _fBestUsedM, DL_LEN_MAX);   // 余料 [m]
iBestA := _iBestACalc;                                            // 最优 A 数量出口 [段]
iBestB := _iBestBCalc;                                            // 最优 B 数量出口 [段]

(* —— 段 7：有效位单点聚合（数量未被截断、原板长度未越域） —— *)
xValid := (iQtyA <= _iQtyAMax) AND (iQtyB <= _iQtyBMax)           // 数量未被钳制截断
          AND (fRibbonLenM <= DL_LEN_MAX)                         // 原板长度未越域
          AND (fOrderLenA > DL_EPS) AND (fOrderLenB > DL_EPS);    // 两种长度均可用
FC_DL_GlassCutOptimizeCalc := xValid;                             // 返回码：TRUE = 计算可信

END_FUNCTION

(* ---- FC_DL_GlassResidualStressCalc.st ---- *)
(*
  Name: FC_DL_GlassResidualStressCalc
  Category: DL_Process
  Version: 1.0.0
  Round: R90 / 2026-11-25
  开源溯源：clean-room 自研（族 浮法玻璃锡槽退火，ST 开源生态实测 0 命中，无外部代码引入）
  功能：1) 残余应力按「温降速率造成的厚度方向温差」估算，逐步为：
             厚度方向温差 ΔT = 温降速率 × 厚度 × 特征均温时间常数
             残余应力 σ = 弹性模量 × 线膨胀系数 × ΔT
           热应力的物理本质是「表面先冷收缩、内部后收缩」，两者收缩量之差受弹性约束即产生应力，
           故应力与「温降速率 × 厚度」成正比，与线膨胀系数、弹性模量成正比。
           特征均温时间常数 DL_TAU_MIN_PER_MM 是「每 mm 厚度对应的热滞后时间」的工程标定值，
           量纲为 min/mm，乘温降速率与厚度后恰好得 °C，不引入额外量纲。
        2) 与安全阈值 DL_SIGMA_SAFE 比较给出 xSafe。退火玻璃的允许残余应力远低于钢化玻璃，
           超阈值意味着切割炸裂与翘曲风险，故上限是硬约束。
  边界条件：1) 非有限值闸：四路实值入参统一过 NOT(x > -DL_BIG AND x < DL_BIG)，
           同时拦 NaN 与 Inf，命中即拦断实值通路（fStressMpa 强制 0.0、xSafe 强制 FALSE）并置无效（R19）。
        2) 分母零闸：本件除数仅为常量，无运行期分母；但三个物性/几何输入都必须为正才具有物理意义，
           故对温降速率、膨胀系数、厚度、弹性模量做 > DL_EPS 的门控（零值判无效）。
        3) 负值闸：温降速率为负（升温）时残余应力符号反转为压应力，本件的判定只面向降温工况，
           故负速率一律判无效而不取绝对值（取绝对值会把升温段误判为有炸裂风险）。
        4) 量程校验：线膨胀系数 0 ~ DL_CTE_MAX(1.0E-4 /°C)、厚度 0 ~ DL_THK_MAX(50 mm)、
           弹性模量 0 ~ DL_E_MAX(300 GPa)、温降速率 0 ~ DL_RATE_MAX(15 °C/min)，越域钳边界但置无效。
        5) 饱和钳制：应力结果钳 0 ~ DL_SIGMA_MAX(1000 MPa)，防组态越界溢出。
  量纲自证：ΔT = (°C/min) × mm × (min/mm) = °C；
           σ = (GPa × 1000 MPa/GPa) × (1/°C) × °C = MPa，量纲闭合；
           1000 为 [MPa/GPa] 弹性模量单位换算因子，无因次混入。
*)

FUNCTION FC_DL_GlassResidualStressCalc : BOOL
VAR_INPUT
    fCoolRateCmin  : REAL;   // 温降速率 [°C/min] / Cooling rate [°C/min]
    fCtePerC       : REAL;   // 线膨胀系数 [1/°C] / Coefficient of thermal expansion [1/°C]
    fThickMm       : REAL;   // 玻璃带厚度 [mm] / Ribbon thickness [mm]
    fYoungGpa      : REAL;   // 弹性模量 [GPa] / Young's modulus [GPa]
END_VAR
VAR_OUTPUT
    fStressMpa     : REAL;   // 估算残余应力 [MPa] / Estimated residual stress [MPa]
    fDeltaTk       : REAL;   // 厚度方向温差（观测用）[°C] / Through-thickness temperature difference [°C]
    xSafe          : BOOL;   // 残余应力安全标志 [bool] / Residual stress safe flag [bool]
    xValid         : BOOL;   // 计算有效标志 [bool] / Calculation valid flag [bool]
END_VAR
VAR
    _fRateClamp    : REAL;   // 钳制后的温降速率 [°C/min] / Clamped cooling rate [°C/min]
    _fThickClamp   : REAL;   // 钳制后的厚度 [mm] / Clamped thickness [mm]
    _fCteClamp     : REAL;   // 钳制后的膨胀系数 [1/°C] / Clamped CTE [1/°C]
    _fYoungClamp   : REAL;   // 钳制后的弹性模量 [GPa] / Clamped Young's modulus [GPa]
    _fDeltaTRaw    : REAL;   // 未饱和的厚度温差 [°C] / Raw through-thickness delta T [°C]
    _fStressRaw    : REAL;   // 未饱和的残余应力 [MPa] / Raw residual stress [MPa]
END_VAR
VAR CONSTANT
    DL_EPS         : REAL := 1.0E-9;    // 零闸阈值 [-] / Zero gate threshold [-]
    DL_BIG         : REAL := 1.0E12;    // 非有限值闸量级上限 [-] / Finiteness gate magnitude [-]
    DL_MPA_PER_GPA : REAL := 1000.0;    // GPa → MPa 换算因子 [MPa/GPa] / Gigapascal to megapascal factor
    DL_TAU_MIN_PER_MM : REAL := 0.50;   // 热滞后时间常数 [min/mm] / Thermal lag time constant [min/mm]
    DL_RATE_MAX    : REAL := 15.0;      // 温降速率量程上限 [°C/min] / Cooling rate range high [°C/min]
    DL_CTE_MAX     : REAL := 1.0E-4;    // 膨胀系数量程上限 [1/°C] / CTE range high [1/°C]
    DL_THK_MAX     : REAL := 50.0;      // 厚度量程上限 [mm] / Thickness range high [mm]
    DL_E_MAX       : REAL := 300.0;     // 弹性模量量程上限 [GPa] / Young's modulus range high [GPa]
    DL_SIGMA_SAFE  : REAL := 7.0;       // 退火残余应力安全阈值 [MPa] / Safe residual stress limit [MPa]
    DL_SIGMA_MAX   : REAL := 1000.0;    // 应力饱和钳制上限 [MPa] / Stress saturation ceiling [MPa]
END_VAR

(* —— 段 1：非有限值闸（R19：四路入参全覆盖，拦 NaN 与 Inf） —— *)
IF NOT (fCoolRateCmin > -DL_BIG AND fCoolRateCmin < DL_BIG)
   OR NOT (fCtePerC > -DL_BIG AND fCtePerC < DL_BIG)
   OR NOT (fThickMm > -DL_BIG AND fThickMm < DL_BIG)
   OR NOT (fYoungGpa > -DL_BIG AND fYoungGpa < DL_BIG) THEN
    fStressMpa := 0.0;                      // 输出强制 0.0 / Output forced to zero
    fDeltaTk := 0.0;                        // 温差强制 0.0 / Delta T forced to zero
    xSafe := FALSE;                         // 安全标志强制 FALSE / Safe flag forced off
    xValid := FALSE;                        // 有效位清零 / Validity cleared
    FC_DL_GlassResidualStressCalc := FALSE; // 返回码同源 / Return mirrors validity
    RETURN;                                 // 立即退出 / Immediate exit
END_IF

(* —— 段 2：零闸与负值闸（物性/几何必须为正；升温工况不属本件判定范围） —— *)
IF (fCoolRateCmin < 0.0) OR (fCtePerC <= DL_EPS) OR (fThickMm <= DL_EPS) OR (fYoungGpa <= DL_EPS) THEN
    fStressMpa := 0.0;                      // 输出强制 0.0 / Output forced to zero
    fDeltaTk := 0.0;                        // 温差强制 0.0 / Delta T forced to zero
    xSafe := FALSE;                         // 安全标志强制 FALSE / Safe flag forced off
    xValid := FALSE;                        // 判无效 / Invalid
    FC_DL_GlassResidualStressCalc := FALSE; // 返回码同步 / Return synchronised
    RETURN;                                 // 提前退出 / Early exit
END_IF

(* —— 段 3：量程钳制（越域钳边界算参考值，段 6 判无效） —— *)
_fRateClamp := LIMIT(0.0, fCoolRateCmin, DL_RATE_MAX);            // 速率钳 0..15 [°C/min]
_fThickClamp := LIMIT(0.0, fThickMm, DL_THK_MAX);                 // 厚度钳 0..50 [mm]
_fCteClamp := LIMIT(0.0, fCtePerC, DL_CTE_MAX);                   // 膨胀系数钳 [1/°C]
_fYoungClamp := LIMIT(0.0, fYoungGpa, DL_E_MAX);                  // 弹性模量钳 [GPa]

(* —— 段 4：厚度温差与残余应力（R22 方向自核：速率与厚度相乘，被时间常数折算为温差） —— *)
_fDeltaTRaw := _fRateClamp * _fThickClamp * DL_TAU_MIN_PER_MM;    // 厚度温差 [°C]
_fStressRaw := _fYoungClamp * DL_MPA_PER_GPA * _fCteClamp * _fDeltaTRaw;   // 残余应力 [MPa]

(* —— 段 5：输出单点写盘（饱和钳制后判安全，保证判据与出口同源） —— *)
fDeltaTk := LIMIT(0.0, _fDeltaTRaw, DL_BIG);                      // 温差出口 [°C]
fStressMpa := LIMIT(0.0, _fStressRaw, DL_SIGMA_MAX);              // 应力出口 [MPa]

(* —— 段 6：有效位单点聚合（四路量程校验） —— *)
xValid := (fCoolRateCmin >= 0.0) AND (fCoolRateCmin <= DL_RATE_MAX)
          AND (fCtePerC > DL_EPS) AND (fCtePerC <= DL_CTE_MAX)
          AND (fThickMm > DL_EPS) AND (fThickMm <= DL_THK_MAX)
          AND (fYoungGpa > DL_EPS) AND (fYoungGpa <= DL_E_MAX);

(* —— 段 7：安全判定（无效数据不得判安全） —— *)
xSafe := xValid AND (fStressMpa <= DL_SIGMA_SAFE);
FC_DL_GlassResidualStressCalc := xValid;                          // 返回码：TRUE = 计算可信

END_FUNCTION

(* ---- FC_DL_GlassRibbonWidthCalc.st ---- *)
(*
  Name: FC_DL_GlassRibbonWidthCalc
  Category: DL_Process
  Version: 1.0.0
  Round: R90 / 2026-11-25
  开源溯源：clean-room 自研（族 浮法玻璃锡槽退火，ST 开源生态实测 0 命中，无外部代码引入）
  功能：1) 玻璃带宽度按「拉边机线速与拉引速度的速度比」投影到目标带宽上估算。
           物理口径：拉边机把玻璃带边缘以 fEdgeRollMps 向外输送，纵向以 fDrawMps 拉引；
           两者相等时带宽维持目标值，比值偏离 1 时带宽按同一比例偏移，
           故 fWidthMm = 目标带宽 × (拉边机线速 / 拉引速度)。
           该式是归一化速度比投影，分子为拉边机线速、分母为拉引速度，方向不可交换
           （交换会得到倒数比，带宽趋势完全反向）。
        2) 与目标带宽比较给出相对偏差 fDevPct = (实测带宽 − 目标带宽) / 目标带宽 × 100，
           正值表示带宽偏宽（拉边过强），负值表示偏窄（拉边不足）。
  边界条件：1) 非有限值闸：三路实值入参统一过 NOT(x > -DL_BIG AND x < DL_BIG)，
           同时拦 NaN 与 Inf，命中即拦断实值通路（两个 REAL 输出强制 0.0）并置无效（R19）。
        2) 分母零闸：ABS(fDrawMps) > DL_EPS（拉引速度为 0 时速度比发散）与
           ABS(fWidthTargetMm) > DL_EPS（目标带宽为 0 时相对偏差无定义）都必须通过，否则判无效。
        3) 负值闸：拉边机线速、拉引速度、目标带宽、容差任一为负判无效
           （速度为负意味着反向运动，不属本件工况，不取绝对值掩盖）。
        4) 速度比窄闸：速度比钳到 DL_SPEED_RATIO_MIN(0.2) ~ DL_SPEED_RATIO_MAX(5.0)，
           越域钳边界算参考值但置无效，防拉引速度极小把带宽放大到无意义量级。
        5) 饱和钳制：带宽结果钳 0 ~ DL_W_MAX_MM(10000 mm)，偏差钳 −1000 ~ +1000 %。
  量纲自证：fWidthMm = mm × (m/s) / (m/s) = mm，速度比无因次，量纲保持长度；
           fDevPct = (mm − mm) / mm × 100 = 无因次 [%]，减法两侧与分母同量纲。
*)

FUNCTION FC_DL_GlassRibbonWidthCalc : BOOL
VAR_INPUT
    fEdgeRollMps   : REAL;   // 拉边机线速度 [m/s] / Edge roller linear speed [m/s]
    fDrawMps       : REAL;   // 玻璃带拉引速度 [m/s] / Ribbon draw speed [m/s]
    fWidthTargetMm : REAL;   // 目标带宽 [mm] / Target ribbon width [mm]
    fTolPct        : REAL;   // 带宽容差（观测用）[%] / Width tolerance for observation [%]
END_VAR
VAR_OUTPUT
    fWidthMm       : REAL;   // 估算带宽 [mm] / Estimated ribbon width [mm]
    fDevPct        : REAL;   // 带宽相对偏差 [%] / Ribbon width relative deviation [%]
    xValid         : BOOL;   // 计算有效标志 [bool] / Calculation valid flag [bool]
END_VAR
VAR
    _fSpeedRatio   : REAL;   // 速度比（拉边 / 拉引）[-] / Speed ratio, edge to draw [-]
    _fWidthRawMm   : REAL;   // 未饱和的带宽 [mm] / Raw ribbon width [mm]
    _fDevRawPct    : REAL;   // 未饱和的偏差 [%] / Raw deviation [%]
END_VAR
VAR CONSTANT
    DL_EPS         : REAL := 1.0E-9;    // 分母零闸阈值 [-] / Division-zero gate threshold [-]
    DL_BIG         : REAL := 1.0E12;    // 非有限值闸量级上限 [-] / Finiteness gate magnitude [-]
    DL_PCT         : REAL := 100.0;     // 百分比换算因子 [%] / Percent conversion factor [%]
    DL_RATIO_MIN   : REAL := 0.20;      // 速度比饱和下限 [-] / Speed ratio saturation low [-]
    DL_RATIO_MAX   : REAL := 5.00;      // 速度比饱和上限 [-] / Speed ratio saturation high [-]
    DL_W_MAX_MM    : REAL := 10000.0;   // 带宽饱和上限 [mm] / Width saturation ceiling [mm]
    DL_DEV_MAX     : REAL := 1000.0;    // 偏差饱和上限 [%] / Deviation saturation ceiling [%]
END_VAR

(* —— 段 1：非有限值闸（R19：四路入参全覆盖，拦 NaN 与 Inf） —— *)
IF NOT (fEdgeRollMps > -DL_BIG AND fEdgeRollMps < DL_BIG)
   OR NOT (fDrawMps > -DL_BIG AND fDrawMps < DL_BIG)
   OR NOT (fWidthTargetMm > -DL_BIG AND fWidthTargetMm < DL_BIG)
   OR NOT (fTolPct > -DL_BIG AND fTolPct < DL_BIG) THEN
    fWidthMm := 0.0;                        // 输出强制 0.0 / Output forced to zero
    fDevPct := 0.0;                         // 偏差强制 0.0 / Deviation forced to zero
    xValid := FALSE;                        // 有效位清零 / Validity cleared
    FC_DL_GlassRibbonWidthCalc := FALSE;    // 返回码同源 / Return mirrors validity
    RETURN;                                 // 立即退出 / Immediate exit
END_IF

(* —— 段 2：分母零闸（R4：拉引速度与目标带宽两个分母） —— *)
IF (ABS(fDrawMps) <= DL_EPS) OR (ABS(fWidthTargetMm) <= DL_EPS) THEN
    fWidthMm := 0.0;                        // 输出强制 0.0 / Output forced to zero
    fDevPct := 0.0;                         // 偏差强制 0.0 / Deviation forced to zero
    xValid := FALSE;                        // 判无效 / Invalid
    FC_DL_GlassRibbonWidthCalc := FALSE;    // 返回码同步 / Return synchronised
    RETURN;                                 // 提前退出 / Early exit
END_IF

(* —— 段 3：负值闸（速度为负意味着反向，不属本工况） —— *)
IF (fEdgeRollMps < 0.0) OR (fDrawMps < 0.0) OR (fWidthTargetMm < 0.0) OR (fTolPct < 0.0) THEN
    fWidthMm := 0.0;                        // 输出强制 0.0 / Output forced to zero
    fDevPct := 0.0;                         // 偏差强制 0.0 / Deviation forced to zero
    xValid := FALSE;                        // 判无效 / Invalid
    FC_DL_GlassRibbonWidthCalc := FALSE;    // 返回码同步 / Return synchronised
    RETURN;                                 // 提前退出 / Early exit
END_IF

(* —— 段 4：速度比归一化（R22 方向自核：拉边机线速在分子、拉引速度在分母） —— *)
_fSpeedRatio := LIMIT(DL_RATIO_MIN, fEdgeRollMps / fDrawMps, DL_RATIO_MAX);   // 速度比 [-]

(* —— 段 5：带宽投影与偏差（分子方向：实测减目标，正值 = 偏宽） —— *)
_fWidthRawMm := fWidthTargetMm * _fSpeedRatio;                    // 带宽 [mm]
_fDevRawPct := (_fWidthRawMm - fWidthTargetMm) / fWidthTargetMm * DL_PCT;   // 偏差 [%]

(* —— 段 6：输出单点写盘（饱和钳制） —— *)
fWidthMm := LIMIT(0.0, _fWidthRawMm, DL_W_MAX_MM);                // 带宽 [mm]
fDevPct := LIMIT(-DL_DEV_MAX, _fDevRawPct, DL_DEV_MAX);           // 偏差 [%]

(* —— 段 7：有效位单点聚合（速度比不越窄闸 + 容差在 0..100 %） —— *)
xValid := (fEdgeRollMps >= 0.0) AND (fDrawMps > DL_EPS)          // 速度为正向
          AND (fWidthTargetMm > DL_EPS)                          // 目标带宽为正
          AND (fTolPct >= 0.0) AND (fTolPct <= DL_PCT)           // 容差在 0..100 %
          AND (fEdgeRollMps / fDrawMps >= DL_RATIO_MIN)          // 速度比不越下限
          AND (fEdgeRollMps / fDrawMps <= DL_RATIO_MAX);         // 速度比不越上限
FC_DL_GlassRibbonWidthCalc := xValid;                            // 返回码：TRUE = 计算可信

END_FUNCTION

(* ---- FC_DL_GlassThicknessCalc.st ---- *)
(*
  Name: FC_DL_GlassThicknessCalc
  Category: DL_Process
  Version: 1.0.0
  Round: R90 / 2026-11-25
  开源溯源：clean-room 自研（族 浮法玻璃锡槽退火，ST 开源生态实测 0 命中，无外部代码引入）
  功能：1) 玻璃带厚度按体积守恒式反算：单位时间流出的玻璃液体积 = 玻璃带截面积 × 拉引速度，
           即 Q = 带宽 × 厚度 × 拉引速度，故厚度 = Q / (带宽 × 拉引速度)。
           全部单位先统一到 SI（m3/s、m、m/s）再计算，最后乘 1000 转 mm；
           不允许混用 m3/h 与 mm 直接相除（那会得到 3.6e6 倍的错误量级）。
        2) 该式是浮法厚度控制的基准式：改厚度只能通过改拉引速度（拉薄/拉厚）或改拉引量实现，
           带宽由拉边机约束，故厚度的可调自由度主要落在速度上。
  边界条件：1) 非有限值闸：三路实值入参统一过 NOT(x > -DL_BIG AND x < DL_BIG)，
           同时拦 NaN 与 Inf，命中即拦断实值通路（fThickMm 强制 0.0）并置无效（R19）。
        2) 分母零闸：带宽按 DL_W_MIN_MM(1.0 mm) 下限钳制后参与除法；
           拉引速度必须 ABS > DL_EPS（速度为 0 表示带不动，厚度无定义），否则判无效。
        3) 负值闸：拉引量、带宽、拉引速度任一为负判无效（不取绝对值掩盖反向）。
        4) 零值语义：拉引量为 0（断板/停拉）时厚度为 0，属合法工况但不具选型意义，
           不判无效；带宽为 0 与速度为 0 判无效（分母不可用）。
        5) 饱和钳制：厚度结果钳 0 ~ DL_THK_MAX_MM(100 mm)，防极小带宽与极低速度组合溢出。
  量纲自证：Q = m3/h ÷ 3600 (s/h) = m3/s；带宽 = mm ÷ 1000 (mm/m) = m；
           Q / (m × m/s) = (m3/s) / (m2/s) = m；再乘 1000 (mm/m) = mm，量纲闭合。
*)

FUNCTION FC_DL_GlassThicknessCalc : BOOL
VAR_INPUT
    fPullM3h       : REAL;   // 玻璃液拉引体积流量 [m3/h] / Glass pull volumetric flow [m3/h]
    fRibbonWidthMm : REAL;   // 玻璃带宽度 [mm] / Ribbon width [mm]
    fDrawMps       : REAL;   // 玻璃带拉引速度 [m/s] / Ribbon draw speed [m/s]
END_VAR
VAR_OUTPUT
    fThickMm       : REAL;   // 玻璃带厚度 [mm] / Ribbon thickness [mm]
    fAreaM2        : REAL;   // 玻璃带截面积（观测用）[m2] / Ribbon cross-section area [m2]
    xValid         : BOOL;   // 计算有效标志 [bool] / Calculation valid flag [bool]
END_VAR
VAR
    _fPullM3s      : REAL;   // 拉引流量 [m3/s] / Pull volumetric flow [m3/s]
    _fWidthM       : REAL;   // 钳制并换算后的带宽 [m] / Clamped width in metres [m]
    _fAreaRawM2    : REAL;   // 截面积 [m2] / Cross-section area [m2]
    _fThickRawM    : REAL;   // 未饱和的厚度 [m] / Raw thickness [m]
END_VAR
VAR CONSTANT
    DL_EPS         : REAL := 1.0E-9;    // 分母零闸阈值 [-] / Division-zero gate threshold [-]
    DL_BIG         : REAL := 1.0E12;    // 非有限值闸量级上限 [-] / Finiteness gate magnitude [-]
    DL_S_PER_H     : REAL := 3600.0;    // h → s 换算因子 [s/h] / Hour to second factor [s/h]
    DL_MM_PER_M    : REAL := 1000.0;    // m → mm 换算因子 [mm/m] / Metre to millimetre factor [mm/m]
    DL_W_MIN_MM    : REAL := 1.0;       // 带宽下限钳制值 [mm] / Width lower clamp [mm]
    DL_THK_MAX_MM  : REAL := 100.0;     // 厚度饱和上限 [mm] / Thickness saturation ceiling [mm]
END_VAR

(* —— 段 1：非有限值闸（R19：三路入参全覆盖，拦 NaN 与 Inf） —— *)
IF NOT (fPullM3h > -DL_BIG AND fPullM3h < DL_BIG)
   OR NOT (fRibbonWidthMm > -DL_BIG AND fRibbonWidthMm < DL_BIG)
   OR NOT (fDrawMps > -DL_BIG AND fDrawMps < DL_BIG) THEN
    fThickMm := 0.0;                        // 输出强制 0.0 / Output forced to zero
    fAreaM2 := 0.0;                         // 截面积强制 0.0 / Area forced to zero
    xValid := FALSE;                        // 有效位清零 / Validity cleared
    FC_DL_GlassThicknessCalc := FALSE;      // 返回码同源 / Return mirrors validity
    RETURN;                                 // 立即退出 / Immediate exit
END_IF

(* —— 段 2：分母零闸（R4：拉引速度是厚度分母） —— *)
IF ABS(fDrawMps) <= DL_EPS THEN
    fThickMm := 0.0;                        // 输出强制 0.0 / Output forced to zero
    fAreaM2 := 0.0;                         // 截面积强制 0.0 / Area forced to zero
    xValid := FALSE;                        // 判无效 / Invalid
    FC_DL_GlassThicknessCalc := FALSE;      // 返回码同步 / Return synchronised
    RETURN;                                 // 提前退出 / Early exit
END_IF

(* —— 段 3：负值闸（流量与几何量均不可为负） —— *)
IF (fPullM3h < 0.0) OR (fRibbonWidthMm < 0.0) OR (fDrawMps < 0.0) THEN
    fThickMm := 0.0;                        // 输出强制 0.0 / Output forced to zero
    fAreaM2 := 0.0;                         // 截面积强制 0.0 / Area forced to zero
    xValid := FALSE;                        // 判无效 / Invalid
    FC_DL_GlassThicknessCalc := FALSE;      // 返回码同步 / Return synchronised
    RETURN;                                 // 提前退出 / Early exit
END_IF

(* —— 段 4：单位统一（m3/h → m3/s，mm → m，两侧都必须先换算） —— *)
_fPullM3s := fPullM3h / DL_S_PER_H;                               // 拉引流量 [m3/s]
_fWidthM := MAX(DL_W_MIN_MM, fRibbonWidthMm) / DL_MM_PER_M;       // 带宽下限钳后换算 [m]

(* —— 段 5：体积守恒主算式（R22 方向自核：流量除以「面积 = 宽 × 速度」） —— *)
_fAreaRawM2 := _fPullM3s / fDrawMps;                              // 截面积 = Q / v [m2]
_fThickRawM := _fAreaRawM2 / _fWidthM;                            // 厚度 = 面积 / 宽 [m]

(* —— 段 6：输出单点写盘（m → mm，饱和钳制） —— *)
fAreaM2 := LIMIT(0.0, _fAreaRawM2, DL_BIG);                       // 截面积 [m2]
fThickMm := LIMIT(0.0, _fThickRawM * DL_MM_PER_M, DL_THK_MAX_MM); // 厚度 [mm]

(* —— 段 7：有效位单点聚合 —— *)
xValid := (fPullM3h >= 0.0)                                       // 拉引量非负
          AND (fRibbonWidthMm >= DL_W_MIN_MM)                     // 带宽不低于下限
          AND (fDrawMps > DL_EPS);                                // 速度为正（分母可用）
FC_DL_GlassThicknessCalc := xValid;                               // 返回码：TRUE = 计算可信

END_FUNCTION

(* ---- FC_DL_GranuleSizeD50Calc.st ---- *)
(*
  DL Factory R84 | FC_DL_GranuleSizeD50Calc
  功能：由累积粒径分布线性插值求 D10/D50/D90 并算跨径距 span
  开源溯源：无（clean-room 自研，依据公开工艺公式，来源=行业通用公式，许可证=MIT，借鉴点=公式结构）
  规则：R1-R16 全遵守
*)
FUNCTION FC_DL_GranuleSizeD50Calc : REAL
VAR_INPUT
    aSizeUm : ARRAY[0..15] OF REAL; // 各档粒径（0..15 号档，单调递增） [µm] / sieve size bins, ascending [um]
    aCumPct : ARRAY[0..15] OF REAL; // 各档累积通过百分比（单调递增） [%] / cumulative passing per bin [%]
    iSampleCnt : INT := 10; // 有效档数（2~16） [档] / effective bin count [bins]
END_VAR
VAR_OUTPUT
    fD10 : REAL; // 10% 通过径 [µm] / size at ten percent passing [um]
    fD90 : REAL; // 90% 通过径 [µm] / size at ninety percent passing [um]
    fSpan : REAL; // 跨径距 (D90−D10)/D50 [-] / span of the distribution [-]
    xValid : BOOL; // 计算结果有效标志 [-] / calculation valid flag [-]
END_VAR
VAR
    i : INT; // 循环游标（1 基起，需访问 i−1 档） [-] / loop cursor starting at one [-]
    fDen : REAL; // 档间累积差（分母，已加下限闸） [%] / inter bin cumulative difference [%]
    fD50 : REAL; // D50 中间量 [µm] / median size intermediate [um]
    xGot10 : BOOL; // 已命中 10% 档标志 [-] / ten percent bin found [-]
    xGot50 : BOOL; // 已命中 50% 档标志 [-] / fifty percent bin found [-]
    xGot90 : BOOL; // 已命中 90% 档标志 [-] / ninety percent bin found [-]
    xFin : BOOL; // 数组有限性判定 [-] / array finiteness verdict [-]
END_VAR

// 段 1｜出口预置（R256）
FC_DL_GranuleSizeD50Calc := -1.0; // 哨兵返回 -1（无效） [-] / sentinel return -1, invalid [-]
fD10 := 0.0; // D10 预置零 [µm] / D10 preset zero [um]
fD90 := 0.0; // D90 预置零 [µm] / D90 preset zero [um]
fSpan := 0.0; // span 预置零 [-] / span preset zero [-]
xValid := FALSE; // 计算完成前不认结果 [-] / unusable before calculation [-]
xGot10 := FALSE; // 命中标志显式清零（FC 局部量不依赖初值） [-] / explicit reset of the hit flag [-]
xGot50 := FALSE; // 命中标志显式清零 [-] / explicit reset of the hit flag [-]
xGot90 := FALSE; // 命中标志显式清零 [-] / explicit reset of the hit flag [-]

// 段 2｜域闸 + 数组有限性闸（R4/R272）
IF iSampleCnt < 2 OR iSampleCnt > 16 THEN
    RETURN; // 少于两档无法插值 [档] / at least two bins needed [bins]
END_IF
xFin := TRUE; // 有限性初值置真 [-] / finiteness starts true [-]
FOR i := 0 TO 15 DO
    IF i < iSampleCnt THEN
        IF NOT (aSizeUm[i] > -1.0E30 AND aSizeUm[i] < 1.0E30) OR NOT (aCumPct[i] > -1.0E30 AND aCumPct[i] < 1.0E30) THEN
            xFin := FALSE; // 任一档非有限即整体无效 [-] / any bad bin voids the result [-]
        END_IF
    END_IF
END_FOR
IF NOT xFin THEN
    RETURN; // 含非有限档值直接退出 [-] / exit on a non finite bin [-]
END_IF

// 段 3｜线性插值定位 D10/D50/D90（首档已越限则直接取首档）
IF aCumPct[0] >= 10.0 THEN
    fD10 := aSizeUm[0]; // 首档已超 10%：D10 取下界 [µm] / first bin above ten percent [um]
    xGot10 := TRUE; // 置命中标志 [-] / mark as found [-]
END_IF
FOR i := 1 TO 15 DO
    IF i < iSampleCnt THEN
        fDen := aCumPct[i] - aCumPct[i - 1]; // % − % = %（档间累积差） / [%] minus [%] = [%]
        IF fDen < 1.0E-9 THEN
            fDen := 1.0E-9; // 分母闸：平台档按极小值兜底，避免除零 [%] / denominator floor [%]
        END_IF
        IF (NOT xGot10) AND (aCumPct[i] >= 10.0) THEN
            fD10 := aSizeUm[i - 1] + ((10.0 - aCumPct[i - 1]) * (aSizeUm[i] - aSizeUm[i - 1])) / fDen; // µm + % × µm ÷ % = µm / [um] + [%] × [um] / [%] = [um]
            xGot10 := TRUE; // 置命中标志 [-] / mark as found [-]
        END_IF
        IF (NOT xGot50) AND (aCumPct[i] >= 50.0) THEN
            fD50 := aSizeUm[i - 1] + ((50.0 - aCumPct[i - 1]) * (aSizeUm[i] - aSizeUm[i - 1])) / fDen; // µm + % × µm ÷ % = µm / [um] + [%] × [um] / [%] = [um]
            xGot50 := TRUE; // 置命中标志 [-] / mark as found [-]
        END_IF
        IF (NOT xGot90) AND (aCumPct[i] >= 90.0) THEN
            fD90 := aSizeUm[i - 1] + ((90.0 - aCumPct[i - 1]) * (aSizeUm[i] - aSizeUm[i - 1])) / fDen; // µm + % × µm ÷ % = µm / [um] + [%] × [um] / [%] = [um]
            xGot90 := TRUE; // 置命中标志 [-] / mark as found [-]
        END_IF
    END_IF
END_FOR
IF (NOT xGot10) OR (NOT xGot50) OR (NOT xGot90) THEN
    RETURN; // 三点未全部命中（分布不完整）拒算 [-] / incomplete distribution rejected [-]
END_IF
IF fD50 < 1.0E-9 THEN
    RETURN; // 分母闸：D50 趋零则 span 无意义 [µm] / denominator gate on D50 [um]
END_IF

// 段 4｜跨径距 span = (D90 − D10) / D50
fSpan := (fD90 - fD10) / fD50; // µm ÷ µm = 无量纲 / [um] / [um] = [-]
IF NOT (fSpan > -1.0E30 AND fSpan < 1.0E30) OR NOT (fD50 > -1.0E30 AND fD50 < 1.0E30) THEN
    RETURN; // 结果非有限再拦一次 [-] / second finiteness gate [-]
END_IF
xValid := TRUE; // 链路有效 [-] / chain valid [-]
FC_DL_GranuleSizeD50Calc := fD50; // 返回 D50 [µm] / return the median size [um]
END_FUNCTION
